  movel([0.304016, -1.350622, -2.573814, -0.787953, 1.570796, 1.874813],accel_mss,speed_ms,0,blend_radius_m)
  movel([0.304007, -1.350886, -2.573637, -0.787866, 1.570796, 1.874804],accel_mss,speed_ms,0,blend_radius_m)
  movel([0.303980, -1.351158, -2.573455, -0.787776, 1.570796, 1.874776],accel_mss,speed_ms,0,blend_radius_m)
  movel([0.303937, -1.351431, -2.573272, -0.787686, 1.570796, 1.874734],accel_mss,speed_ms,0,blend_radius_m)
  movel([0.303879, -1.351709, -2.573085, -0.787594, 1.570796, 1.874675],accel_mss,speed_ms,0,blend_radius_m)
  movel([0.303801, -1.351990, -2.572896, -0.787502, 1.570796, 1.874598],accel_mss,speed_ms,0,blend_radius_m)
  movel([0.303710, -1.352271, -2.572708, -0.787410, 1.570796, 1.874506],accel_mss,speed_ms,0,blend_radius_m)
  movel([0.303601, -1.352553, -2.572519, -0.787318, 1.570796, 1.874397],accel_mss,speed_ms,0,blend_radius_m)
  movel([0.303476, -1.352836, -2.572328, -0.787225, 1.570796, 1.874272],accel_mss,speed_ms,0,blend_radius_m)
  movel([0.303336, -1.353119, -2.572138, -0.787132, 1.570796, 1.874133],accel_mss,speed_ms,0,blend_radius_m)
  movel([0.303181, -1.353399, -2.571949, -0.787041, 1.570796, 1.873978],accel_mss,speed_ms,0,blend_radius_m)
  movel([0.303018, -1.353668, -2.571768, -0.786953, 1.570796, 1.873815],accel_mss,speed_ms,0,blend_radius_m)
  movel([0.302839, -1.353937, -2.571586, -0.786865, 1.570796, 1.873636],accel_mss,speed_ms,0,blend_radius_m)
  movel([0.302653, -1.354200, -2.571409, -0.786780, 1.570796, 1.873449],accel_mss,speed_ms,0,blend_radius_m)
  movel([0.302453, -1.354460, -2.571234, -0.786695, 1.570796, 1.873250],accel_mss,speed_ms,0,blend_radius_m)
  movel([0.302246, -1.354707, -2.571067, -0.786615, 1.570796, 1.873043],accel_mss,speed_ms,0,blend_radius_m)
  movel([0.302029, -1.354951, -2.570903, -0.786536, 1.570796, 1.872825],accel_mss,speed_ms,0,blend_radius_m)
  movel([0.301802, -1.355186, -2.570743, -0.786459, 1.570796, 1.872599],accel_mss,speed_ms,0,blend_radius_m)
  movel([0.301564, -1.355414, -2.570589, -0.786386, 1.570796, 1.872361],accel_mss,speed_ms,0,blend_radius_m)
  movel([0.301323, -1.355631, -2.570442, -0.786315, 1.570796, 1.872119],accel_mss,speed_ms,0,blend_radius_m)
  movel([0.301073, -1.355840, -2.570301, -0.786248, 1.570796, 1.871869],accel_mss,speed_ms,0,blend_radius_m)
  movel([0.300816, -1.356039, -2.570167, -0.786184, 1.570796, 1.871613],accel_mss,speed_ms,0,blend_radius_m)
  movel([0.300551, -1.356229, -2.570038, -0.786122, 1.570796, 1.871347],accel_mss,speed_ms,0,blend_radius_m)
  movel([0.300280, -1.356409, -2.569916, -0.786064, 1.570796, 1.871076],accel_mss,speed_ms,0,blend_radius_m)
  movel([0.300006, -1.356576, -2.569803, -0.786010, 1.570796, 1.870802],accel_mss,speed_ms,0,blend_radius_m)
  movel([0.299729, -1.356732, -2.569697, -0.785960, 1.570796, 1.870525],accel_mss,speed_ms,0,blend_radius_m)
  movel([0.299446, -1.356878, -2.569598, -0.785913, 1.570796, 1.870242],accel_mss,speed_ms,0,blend_radius_m)
  movel([0.299211, -1.356989, -2.569523, -0.785877, 1.570796, 1.870008],accel_mss,speed_ms,0,blend_radius_m)
  movel([0.298976, -1.357089, -2.569455, -0.785845, 1.570796, 1.869772],accel_mss,speed_ms,0,blend_radius_m)
  movel([0.298781, -1.357162, -2.569405, -0.785822, 1.570796, 1.869578],accel_mss,speed_ms,0,blend_radius_m)
  movel([0.298590, -1.357219, -2.569366, -0.785803, 1.570796, 1.869386],accel_mss,speed_ms,0,blend_radius_m)
  movel([0.298374, -1.357273, -2.569330, -0.785786, 1.570796, 1.869170],accel_mss,speed_ms,0,blend_radius_m)
  movel([0.298159, -1.357310, -2.569305, -0.785774, 1.570796, 1.868955],accel_mss,speed_ms,0,blend_radius_m)
  movel([0.297828, -1.357357, -2.569273, -0.785759, 1.570796, 1.868625],accel_mss,speed_ms,0,blend_radius_m)
  movel([0.297500, -1.357396, -2.569246, -0.785747, 1.570796, 1.868297],accel_mss,speed_ms,0,blend_radius_m)
  movel([0.297176, -1.357431, -2.569223, -0.785735, 1.570796, 1.867972],accel_mss,speed_ms,0,blend_radius_m)
  movel([0.296852, -1.357459, -2.569204, -0.785726, 1.570796, 1.867648],accel_mss,speed_ms,0,blend_radius_m)
  movel([0.296645, -1.357469, -2.569197, -0.785723, 1.570796, 1.867441],accel_mss,speed_ms,0,blend_radius_m)
  movel([0.296449, -1.357463, -2.569201, -0.785725, 1.570796, 1.867245],accel_mss,speed_ms,0,blend_radius_m)
  movel([0.296278, -1.357446, -2.569212, -0.785730, 1.570796, 1.867075],accel_mss,speed_ms,0,blend_radius_m)
  movel([0.296121, -1.357413, -2.569235, -0.785741, 1.570796, 1.866917],accel_mss,speed_ms,0,blend_radius_m)
  movel([0.295935, -1.357359, -2.569272, -0.785759, 1.570796, 1.866731],accel_mss,speed_ms,0,blend_radius_m)
  movel([0.295754, -1.357297, -2.569313, -0.785778, 1.570796, 1.866550],accel_mss,speed_ms,0,blend_radius_m)
  movel([0.295553, -1.357209, -2.569373, -0.785807, 1.570796, 1.866349],accel_mss,speed_ms,0,blend_radius_m)
  movel([0.295368, -1.357105, -2.569444, -0.785840, 1.570796, 1.866165],accel_mss,speed_ms,0,blend_radius_m)
  movel([0.295196, -1.356987, -2.569524, -0.785878, 1.570796, 1.865992],accel_mss,speed_ms,0,blend_radius_m)
  movel([0.295024, -1.356844, -2.569621, -0.785924, 1.570796, 1.865820],accel_mss,speed_ms,0,blend_radius_m)
  movel([0.294865, -1.356689, -2.569726, -0.785974, 1.570796, 1.865661],accel_mss,speed_ms,0,blend_radius_m)
  movel([0.294721, -1.356523, -2.569839, -0.786028, 1.570796, 1.865518],accel_mss,speed_ms,0,blend_radius_m)
  movel([0.294587, -1.356342, -2.569961, -0.786086, 1.570796, 1.865383],accel_mss,speed_ms,0,blend_radius_m)
  movel([0.294469, -1.356148, -2.570092, -0.786148, 1.570796, 1.865265],accel_mss,speed_ms,0,blend_radius_m)
  movel([0.294364, -1.355946, -2.570229, -0.786214, 1.570796, 1.865161],accel_mss,speed_ms,0,blend_radius_m)
  movel([0.294280, -1.355740, -2.570369, -0.786280, 1.570796, 1.865076],accel_mss,speed_ms,0,blend_radius_m)
  movel([0.294210, -1.355524, -2.570515, -0.786350, 1.570796, 1.865007],accel_mss,speed_ms,0,blend_radius_m)
  movel([0.294158, -1.355298, -2.570668, -0.786423, 1.570796, 1.864954],accel_mss,speed_ms,0,blend_radius_m)
  movel([0.294120, -1.355064, -2.570826, -0.786499, 1.570796, 1.864916],accel_mss,speed_ms,0,blend_radius_m)
  movel([0.294091, -1.354823, -2.570988, -0.786577, 1.570796, 1.864887],accel_mss,speed_ms,0,blend_radius_m)
  movel([0.294085, -1.354708, -2.571067, -0.786615, 1.570796, 1.864882],accel_mss,speed_ms,0,blend_radius_m)
  movel([0.294088, -1.354589, -2.571147, -0.786653, 1.570796, 1.864884],accel_mss,speed_ms,0,blend_radius_m)
  movel([0.294101, -1.354467, -2.571229, -0.786693, 1.570796, 1.864897],accel_mss,speed_ms,0,blend_radius_m)
  movel([0.294142, -1.354249, -2.571376, -0.786764, 1.570796, 1.864938],accel_mss,speed_ms,0,blend_radius_m)
  movel([0.294198, -1.354028, -2.571525, -0.786836, 1.570796, 1.864995],accel_mss,speed_ms,0,blend_radius_m)
  speed_ms = 0.003
  movel([0.294198, -1.341397, -2.565271, -0.805721, 1.570796, 1.864995],accel_mss,speed_ms,0,blend_radius_m)
  speed_ms = 0.01
  movel([0.294198, -1.317224, -2.552384, -0.842780, 1.570796, 1.864995],accel_mss,speed_ms,0,blend_radius_m)
  movel([0.288042, -1.339808, -2.537610, -0.834971, 1.570796, 1.858839],accel_mss,speed_ms,0,blend_radius_m)
  movel([0.288042, -1.363639, -2.550213, -0.798536, 1.570796, 1.858839],accel_mss,speed_ms,0,blend_radius_m)
  speed_ms = 0.003
  movel([0.288042, -1.372930, -2.554809, -0.784650, 1.570796, 1.858839],accel_mss,speed_ms,0,blend_radius_m)
  speed_ms = 0.007
  movel([0.288122, -1.372941, -2.554802, -0.784647, 1.570796, 1.858918],accel_mss,speed_ms,0,blend_radius_m)
  movel([0.288195, -1.372963, -2.554786, -0.784640, 1.570796, 1.858991],accel_mss,speed_ms,0,blend_radius_m)
  movel([0.288260, -1.372997, -2.554762, -0.784630, 1.570796, 1.859056],accel_mss,speed_ms,0,blend_radius_m)
  movel([0.288326, -1.373050, -2.554725, -0.784614, 1.570796, 1.859122],accel_mss,speed_ms,0,blend_radius_m)
  movel([0.288376, -1.373118, -2.554677, -0.784594, 1.570796, 1.859172],accel_mss,speed_ms,0,blend_radius_m)
  movel([0.288408, -1.373199, -2.554620, -0.784569, 1.570796, 1.859204],accel_mss,speed_ms,0,blend_radius_m)
  movel([0.288418, -1.373289, -2.554557, -0.784543, 1.570796, 1.859215],accel_mss,speed_ms,0,blend_radius_m)
  movel([0.288412, -1.373390, -2.554486, -0.784513, 1.570796, 1.859208],accel_mss,speed_ms,0,blend_radius_m)
  movel([0.288388, -1.373495, -2.554413, -0.784482, 1.570796, 1.859185],accel_mss,speed_ms,0,blend_radius_m)
  movel([0.288346, -1.373602, -2.554338, -0.784450, 1.570796, 1.859142],accel_mss,speed_ms,0,blend_radius_m)
  movel([0.288285, -1.373708, -2.554263, -0.784418, 1.570796, 1.859081],accel_mss,speed_ms,0,blend_radius_m)
  movel([0.288212, -1.373810, -2.554191, -0.784388, 1.570796, 1.859008],accel_mss,speed_ms,0,blend_radius_m)
  movel([0.288127, -1.373904, -2.554125, -0.784360, 1.570796, 1.858924],accel_mss,speed_ms,0,blend_radius_m)
  movel([0.288029, -1.373991, -2.554064, -0.784334, 1.570796, 1.858825],accel_mss,speed_ms,0,blend_radius_m)
  movel([0.287923, -1.374066, -2.554011, -0.784312, 1.570796, 1.858720],accel_mss,speed_ms,0,blend_radius_m)
  movel([0.287837, -1.374115, -2.553977, -0.784297, 1.570796, 1.858633],accel_mss,speed_ms,0,blend_radius_m)
  movel([0.287749, -1.374155, -2.553948, -0.784285, 1.570796, 1.858545],accel_mss,speed_ms,0,blend_radius_m)
  movel([0.287660, -1.374183, -2.553929, -0.784277, 1.570796, 1.858456],accel_mss,speed_ms,0,blend_radius_m)
  movel([0.287572, -1.374202, -2.553916, -0.784272, 1.570796, 1.858368],accel_mss,speed_ms,0,blend_radius_m)
  movel([0.287487, -1.374207, -2.553912, -0.784270, 1.570796, 1.858284],accel_mss,speed_ms,0,blend_radius_m)
  movel([0.287398, -1.374200, -2.553917, -0.784272, 1.570796, 1.858194],accel_mss,speed_ms,0,blend_radius_m)
  movel([0.287321, -1.374176, -2.553934, -0.784279, 1.570796, 1.858117],accel_mss,speed_ms,0,blend_radius_m)
  movel([0.287255, -1.374136, -2.553962, -0.784291, 1.570796, 1.858052],accel_mss,speed_ms,0,blend_radius_m)
  movel([0.287198, -1.374077, -2.554003, -0.784308, 1.570796, 1.857994],accel_mss,speed_ms,0,blend_radius_m)
  movel([0.287153, -1.374009, -2.554052, -0.784329, 1.570796, 1.857949],accel_mss,speed_ms,0,blend_radius_m)
  movel([0.287124, -1.373932, -2.554106, -0.784352, 1.570796, 1.857921],accel_mss,speed_ms,0,blend_radius_m)
  movel([0.287110, -1.373847, -2.554166, -0.784377, 1.570796, 1.857906],accel_mss,speed_ms,0,blend_radius_m)
  movel([0.287111, -1.373755, -2.554230, -0.784404, 1.570796, 1.857907],accel_mss,speed_ms,0,blend_radius_m)
  movel([0.287127, -1.373658, -2.554298, -0.784433, 1.570796, 1.857924],accel_mss,speed_ms,0,blend_radius_m)
  movel([0.287155, -1.373568, -2.554361, -0.784460, 1.570796, 1.857952],accel_mss,speed_ms,0,blend_radius_m)
  movel([0.287204, -1.373478, -2.554425, -0.784487, 1.570796, 1.858000],accel_mss,speed_ms,0,blend_radius_m)
  movel([0.287266, -1.373390, -2.554486, -0.784513, 1.570796, 1.858062],accel_mss,speed_ms,0,blend_radius_m)
  movel([0.287346, -1.373301, -2.554549, -0.784539, 1.570796, 1.858143],accel_mss,speed_ms,0,blend_radius_m)
  movel([0.287430, -1.373215, -2.554609, -0.784565, 1.570796, 1.858227],accel_mss,speed_ms,0,blend_radius_m)
  movel([0.287524, -1.373135, -2.554665, -0.784589, 1.570796, 1.858321],accel_mss,speed_ms,0,blend_radius_m)
  movel([0.287608, -1.373073, -2.554709, -0.784607, 1.570796, 1.858404],accel_mss,speed_ms,0,blend_radius_m)
  movel([0.287698, -1.373019, -2.554746, -0.784623, 1.570796, 1.858494],accel_mss,speed_ms,0,blend_radius_m)
  movel([0.287789, -1.372976, -2.554777, -0.784636, 1.570796, 1.858586],accel_mss,speed_ms,0,blend_radius_m)
  movel([0.287876, -1.372949, -2.554796, -0.784644, 1.570796, 1.858672],accel_mss,speed_ms,0,blend_radius_m)
  movel([0.287961, -1.372933, -2.554807, -0.784649, 1.570796, 1.858758],accel_mss,speed_ms,0,blend_radius_m)
  movel([0.288042, -1.372930, -2.554809, -0.784650, 1.570796, 1.858839],accel_mss,speed_ms,0,blend_radius_m)
  speed_ms = 0.003
  movel([0.288042, -1.376070, -2.556325, -0.779994, 1.570796, 1.858839],accel_mss,speed_ms,0,blend_radius_m)
  speed_ms = 0.007
  movel([0.288122, -1.376081, -2.556317, -0.779991, 1.570796, 1.858918],accel_mss,speed_ms,0,blend_radius_m)
  movel([0.288195, -1.376103, -2.556302, -0.779984, 1.570796, 1.858991],accel_mss,speed_ms,0,blend_radius_m)
  movel([0.288260, -1.376137, -2.556278, -0.779974, 1.570796, 1.859056],accel_mss,speed_ms,0,blend_radius_m)
  movel([0.288326, -1.376190, -2.556241, -0.779958, 1.570796, 1.859122],accel_mss,speed_ms,0,blend_radius_m)
  movel([0.288376, -1.376258, -2.556193, -0.779938, 1.570796, 1.859172],accel_mss,speed_ms,0,blend_radius_m)
  movel([0.288408, -1.376339, -2.556136, -0.779915, 1.570796, 1.859204],accel_mss,speed_ms,0,blend_radius_m)
  movel([0.288418, -1.376429, -2.556072, -0.779888, 1.570796, 1.859215],accel_mss,speed_ms,0,blend_radius_m)
  movel([0.288412, -1.376529, -2.556001, -0.779859, 1.570796, 1.859208],accel_mss,speed_ms,0,blend_radius_m)
  movel([0.288388, -1.376634, -2.555928, -0.779828, 1.570796, 1.859185],accel_mss,speed_ms,0,blend_radius_m)
  movel([0.288346, -1.376740, -2.555852, -0.779796, 1.570796, 1.859142],accel_mss,speed_ms,0,blend_radius_m)
  movel([0.288285, -1.376847, -2.555777, -0.779765, 1.570796, 1.859081],accel_mss,speed_ms,0,blend_radius_m)
  movel([0.288212, -1.376948, -2.555706, -0.779735, 1.570796, 1.859008],accel_mss,speed_ms,0,blend_radius_m)
  movel([0.288127, -1.377042, -2.555639, -0.779708, 1.570796, 1.858924],accel_mss,speed_ms,0,blend_radius_m)
  movel([0.288029, -1.377129, -2.555578, -0.779682, 1.570796, 1.858825],accel_mss,speed_ms,0,blend_radius_m)
  movel([0.287923, -1.377204, -2.555525, -0.779660, 1.570796, 1.858720],accel_mss,speed_ms,0,blend_radius_m)
  movel([0.287837, -1.377252, -2.555491, -0.779646, 1.570796, 1.858633],accel_mss,speed_ms,0,blend_radius_m)
  movel([0.287749, -1.377293, -2.555462, -0.779634, 1.570796, 1.858545],accel_mss,speed_ms,0,blend_radius_m)
  movel([0.287660, -1.377320, -2.555443, -0.779626, 1.570796, 1.858456],accel_mss,speed_ms,0,blend_radius_m)
  movel([0.287572, -1.377339, -2.555430, -0.779621, 1.570796, 1.858368],accel_mss,speed_ms,0,blend_radius_m)
  movel([0.287487, -1.377344, -2.555426, -0.779619, 1.570796, 1.858284],accel_mss,speed_ms,0,blend_radius_m)
  movel([0.287398, -1.377337, -2.555431, -0.779621, 1.570796, 1.858194],accel_mss,speed_ms,0,blend_radius_m)
  movel([0.287321, -1.377313, -2.555448, -0.779628, 1.570796, 1.858117],accel_mss,speed_ms,0,blend_radius_m)
  movel([0.287255, -1.377273, -2.555476, -0.779640, 1.570796, 1.858052],accel_mss,speed_ms,0,blend_radius_m)
  movel([0.287198, -1.377215, -2.555517, -0.779657, 1.570796, 1.857994],accel_mss,speed_ms,0,blend_radius_m)
  movel([0.287153, -1.377146, -2.555566, -0.779677, 1.570796, 1.857949],accel_mss,speed_ms,0,blend_radius_m)
  movel([0.287124, -1.377069, -2.555620, -0.779700, 1.570796, 1.857921],accel_mss,speed_ms,0,blend_radius_m)
  movel([0.287110, -1.376985, -2.555680, -0.779725, 1.570796, 1.857906],accel_mss,speed_ms,0,blend_radius_m)
  movel([0.287111, -1.376894, -2.555744, -0.779751, 1.570796, 1.857907],accel_mss,speed_ms,0,blend_radius_m)
  movel([0.287127, -1.376796, -2.555813, -0.779780, 1.570796, 1.857924],accel_mss,speed_ms,0,blend_radius_m)
  movel([0.287155, -1.376707, -2.555876, -0.779806, 1.570796, 1.857952],accel_mss,speed_ms,0,blend_radius_m)
  movel([0.287204, -1.376617, -2.555940, -0.779833, 1.570796, 1.858000],accel_mss,speed_ms,0,blend_radius_m)
  movel([0.287266, -1.376529, -2.556001, -0.779858, 1.570796, 1.858062],accel_mss,speed_ms,0,blend_radius_m)
  movel([0.287346, -1.376440, -2.556064, -0.779885, 1.570796, 1.858143],accel_mss,speed_ms,0,blend_radius_m)
  movel([0.287430, -1.376355, -2.556124, -0.779910, 1.570796, 1.858227],accel_mss,speed_ms,0,blend_radius_m)
  movel([0.287524, -1.376275, -2.556181, -0.779933, 1.570796, 1.858321],accel_mss,speed_ms,0,blend_radius_m)
  movel([0.287608, -1.376213, -2.556224, -0.779952, 1.570796, 1.858404],accel_mss,speed_ms,0,blend_radius_m)
  movel([0.287698, -1.376160, -2.556262, -0.779967, 1.570796, 1.858494],accel_mss,speed_ms,0,blend_radius_m)
  movel([0.287789, -1.376117, -2.556292, -0.779980, 1.570796, 1.858586],accel_mss,speed_ms,0,blend_radius_m)
  movel([0.287876, -1.376089, -2.556311, -0.779988, 1.570796, 1.858672],accel_mss,speed_ms,0,blend_radius_m)
  movel([0.287961, -1.376073, -2.556323, -0.779993, 1.570796, 1.858758],accel_mss,speed_ms,0,blend_radius_m)
  movel([0.288042, -1.376070, -2.556325, -0.779994, 1.570796, 1.858839],accel_mss,speed_ms,0,blend_radius_m)
  speed_ms = 0.003
  movel([0.288042, -1.363639, -2.550213, -0.798536, 1.570796, 1.858839],accel_mss,speed_ms,0,blend_radius_m)
  speed_ms = 0.01
  movel([0.288042, -1.339808, -2.537610, -0.834971, 1.570796, 1.858839],accel_mss,speed_ms,0,blend_radius_m)
  movel([0.266011, -1.335427, -2.540528, -0.836434, 1.570796, 1.836807],accel_mss,speed_ms,0,blend_radius_m)
  movel([0.266011, -1.359326, -2.553186, -0.799877, 1.570796, 1.836807],accel_mss,speed_ms,0,blend_radius_m)
  speed_ms = 0.003
  movel([0.266011, -1.368646, -2.557802, -0.785941, 1.570796, 1.836807],accel_mss,speed_ms,0,blend_radius_m)
  speed_ms = 0.007
  movel([0.265722, -1.369059, -2.557515, -0.785815, 1.570796, 1.836519],accel_mss,speed_ms,0,blend_radius_m)
  movel([0.265423, -1.369470, -2.557229, -0.785690, 1.570796, 1.836219],accel_mss,speed_ms,0,blend_radius_m)
  movel([0.265112, -1.369875, -2.556947, -0.785568, 1.570796, 1.835909],accel_mss,speed_ms,0,blend_radius_m)
  movel([0.264791, -1.370276, -2.556667, -0.785446, 1.570796, 1.835587],accel_mss,speed_ms,0,blend_radius_m)
  movel([0.264465, -1.370663, -2.556397, -0.785330, 1.570796, 1.835261],accel_mss,speed_ms,0,blend_radius_m)
  movel([0.264126, -1.371044, -2.556130, -0.785215, 1.570796, 1.834923],accel_mss,speed_ms,0,blend_radius_m)
  movel([0.263781, -1.371418, -2.555869, -0.785102, 1.570796, 1.834578],accel_mss,speed_ms,0,blend_radius_m)
  movel([0.263424, -1.371787, -2.555611, -0.784992, 1.570796, 1.834220],accel_mss,speed_ms,0,blend_radius_m)
  movel([0.263058, -1.372146, -2.555359, -0.784884, 1.570796, 1.833855],accel_mss,speed_ms,0,blend_radius_m)
  movel([0.262685, -1.372499, -2.555111, -0.784778, 1.570796, 1.833481],accel_mss,speed_ms,0,blend_radius_m)
  movel([0.262301, -1.372843, -2.554870, -0.784676, 1.570796, 1.833097],accel_mss,speed_ms,0,blend_radius_m)
  movel([0.261910, -1.373179, -2.554634, -0.784575, 1.570796, 1.832707],accel_mss,speed_ms,0,blend_radius_m)
  movel([0.261537, -1.373487, -2.554418, -0.784484, 1.570796, 1.832333],accel_mss,speed_ms,0,blend_radius_m)
  movel([0.261156, -1.373790, -2.554205, -0.784394, 1.570796, 1.831952],accel_mss,speed_ms,0,blend_radius_m)
  movel([0.260769, -1.374082, -2.554000, -0.784307, 1.570796, 1.831565],accel_mss,speed_ms,0,blend_radius_m)
  movel([0.260377, -1.374369, -2.553798, -0.784222, 1.570796, 1.831173],accel_mss,speed_ms,0,blend_radius_m)
  movel([0.259998, -1.374634, -2.553611, -0.784143, 1.570796, 1.830795],accel_mss,speed_ms,0,blend_radius_m)
  movel([0.259613, -1.374890, -2.553431, -0.784068, 1.570796, 1.830409],accel_mss,speed_ms,0,blend_radius_m)
  movel([0.259224, -1.375137, -2.553257, -0.783995, 1.570796, 1.830020],accel_mss,speed_ms,0,blend_radius_m)
  movel([0.258830, -1.375375, -2.553090, -0.783925, 1.570796, 1.829626],accel_mss,speed_ms,0,blend_radius_m)
  movel([0.258430, -1.375602, -2.552929, -0.783858, 1.570796, 1.829227],accel_mss,speed_ms,0,blend_radius_m)
  movel([0.258032, -1.375819, -2.552776, -0.783794, 1.570796, 1.828828],accel_mss,speed_ms,0,blend_radius_m)
  movel([0.257627, -1.376026, -2.552630, -0.783733, 1.570796, 1.828423],accel_mss,speed_ms,0,blend_radius_m)
  movel([0.257223, -1.376222, -2.552492, -0.783675, 1.570796, 1.828019],accel_mss,speed_ms,0,blend_radius_m)
  movel([0.256797, -1.376415, -2.552356, -0.783619, 1.570796, 1.827593],accel_mss,speed_ms,0,blend_radius_m)
  movel([0.256368, -1.376599, -2.552225, -0.783565, 1.570796, 1.827165],accel_mss,speed_ms,0,blend_radius_m)
  movel([0.255939, -1.376774, -2.552102, -0.783514, 1.570796, 1.826735],accel_mss,speed_ms,0,blend_radius_m)
  movel([0.255510, -1.376937, -2.551986, -0.783466, 1.570796, 1.826306],accel_mss,speed_ms,0,blend_radius_m)
  movel([0.255204, -1.377044, -2.551910, -0.783434, 1.570796, 1.826001],accel_mss,speed_ms,0,blend_radius_m)
  movel([0.254900, -1.377139, -2.551843, -0.783407, 1.570796, 1.825697],accel_mss,speed_ms,0,blend_radius_m)
  movel([0.254597, -1.377223, -2.551784, -0.783382, 1.570796, 1.825393],accel_mss,speed_ms,0,blend_radius_m)
  movel([0.254295, -1.377294, -2.551734, -0.783361, 1.570796, 1.825092],accel_mss,speed_ms,0,blend_radius_m)
  movel([0.253772, -1.377400, -2.551658, -0.783330, 1.570796, 1.824569],accel_mss,speed_ms,0,blend_radius_m)
  movel([0.253251, -1.377494, -2.551592, -0.783303, 1.570796, 1.824047],accel_mss,speed_ms,0,blend_radius_m)
  movel([0.252731, -1.377575, -2.551535, -0.783279, 1.570796, 1.823527],accel_mss,speed_ms,0,blend_radius_m)
  movel([0.252217, -1.377643, -2.551487, -0.783259, 1.570796, 1.823013],accel_mss,speed_ms,0,blend_radius_m)
  movel([0.251706, -1.377697, -2.551448, -0.783244, 1.570796, 1.822503],accel_mss,speed_ms,0,blend_radius_m)
  movel([0.251202, -1.377738, -2.551419, -0.783232, 1.570796, 1.821998],accel_mss,speed_ms,0,blend_radius_m)
  movel([0.250916, -1.377752, -2.551409, -0.783228, 1.570796, 1.821712],accel_mss,speed_ms,0,blend_radius_m)
  movel([0.250636, -1.377752, -2.551409, -0.783228, 1.570796, 1.821432],accel_mss,speed_ms,0,blend_radius_m)
  movel([0.250362, -1.377741, -2.551417, -0.783231, 1.570796, 1.821158],accel_mss,speed_ms,0,blend_radius_m)
  movel([0.250093, -1.377716, -2.551435, -0.783238, 1.570796, 1.820890],accel_mss,speed_ms,0,blend_radius_m)
  movel([0.249712, -1.377667, -2.551469, -0.783252, 1.570796, 1.820508],accel_mss,speed_ms,0,blend_radius_m)
  movel([0.249339, -1.377604, -2.551514, -0.783271, 1.570796, 1.820135],accel_mss,speed_ms,0,blend_radius_m)
  movel([0.248973, -1.377532, -2.551565, -0.783292, 1.570796, 1.819770],accel_mss,speed_ms,0,blend_radius_m)
  movel([0.248614, -1.377446, -2.551626, -0.783317, 1.570796, 1.819410],accel_mss,speed_ms,0,blend_radius_m)
  movel([0.248285, -1.377354, -2.551691, -0.783344, 1.570796, 1.819082],accel_mss,speed_ms,0,blend_radius_m)
  movel([0.247963, -1.377248, -2.551766, -0.783375, 1.570796, 1.818759],accel_mss,speed_ms,0,blend_radius_m)
  movel([0.247652, -1.377131, -2.551849, -0.783409, 1.570796, 1.818449],accel_mss,speed_ms,0,blend_radius_m)
  movel([0.247353, -1.376999, -2.551943, -0.783448, 1.570796, 1.818149],accel_mss,speed_ms,0,blend_radius_m)
  movel([0.247061, -1.376856, -2.552043, -0.783489, 1.570796, 1.817857],accel_mss,speed_ms,0,blend_radius_m)
  movel([0.246782, -1.376699, -2.552154, -0.783535, 1.570796, 1.817578],accel_mss,speed_ms,0,blend_radius_m)
  movel([0.246513, -1.376530, -2.552274, -0.783585, 1.570796, 1.817309],accel_mss,speed_ms,0,blend_radius_m)
  movel([0.246253, -1.376351, -2.552401, -0.783637, 1.570796, 1.817050],accel_mss,speed_ms,0,blend_radius_m)
  movel([0.245991, -1.376146, -2.552545, -0.783697, 1.570796, 1.816788],accel_mss,speed_ms,0,blend_radius_m)
  movel([0.245739, -1.375930, -2.552698, -0.783761, 1.570796, 1.816536],accel_mss,speed_ms,0,blend_radius_m)
  movel([0.245496, -1.375706, -2.552856, -0.783827, 1.570796, 1.816292],accel_mss,speed_ms,0,blend_radius_m)
  movel([0.245264, -1.375473, -2.553020, -0.783896, 1.570796, 1.816060],accel_mss,speed_ms,0,blend_radius_m)
  movel([0.245040, -1.375220, -2.553198, -0.783970, 1.570796, 1.815836],accel_mss,speed_ms,0,blend_radius_m)
  movel([0.244827, -1.374957, -2.553384, -0.784048, 1.570796, 1.815624],accel_mss,speed_ms,0,blend_radius_m)
  movel([0.244629, -1.374686, -2.553575, -0.784128, 1.570796, 1.815425],accel_mss,speed_ms,0,blend_radius_m)
  movel([0.244442, -1.374403, -2.553774, -0.784212, 1.570796, 1.815238],accel_mss,speed_ms,0,blend_radius_m)
  movel([0.244275, -1.374114, -2.553978, -0.784298, 1.570796, 1.815071],accel_mss,speed_ms,0,blend_radius_m)
  movel([0.244119, -1.373818, -2.554185, -0.784385, 1.570796, 1.814915],accel_mss,speed_ms,0,blend_radius_m)
  movel([0.243980, -1.373509, -2.554403, -0.784477, 1.570796, 1.814777],accel_mss,speed_ms,0,blend_radius_m)
  movel([0.243857, -1.373194, -2.554624, -0.784571, 1.570796, 1.814654],accel_mss,speed_ms,0,blend_radius_m)
  movel([0.243743, -1.372861, -2.554857, -0.784670, 1.570796, 1.814539],accel_mss,speed_ms,0,blend_radius_m)
  movel([0.243647, -1.372520, -2.555097, -0.784772, 1.570796, 1.814444],accel_mss,speed_ms,0,blend_radius_m)
  movel([0.243565, -1.372169, -2.555343, -0.784877, 1.570796, 1.814362],accel_mss,speed_ms,0,blend_radius_m)
  movel([0.243497, -1.371812, -2.555593, -0.784984, 1.570796, 1.814293],accel_mss,speed_ms,0,blend_radius_m)
  movel([0.243441, -1.371423, -2.555865, -0.785101, 1.570796, 1.814237],accel_mss,speed_ms,0,blend_radius_m)
  movel([0.243401, -1.371029, -2.556141, -0.785219, 1.570796, 1.814197],accel_mss,speed_ms,0,blend_radius_m)
  movel([0.243370, -1.370631, -2.556418, -0.785339, 1.570796, 1.814167],accel_mss,speed_ms,0,blend_radius_m)
  movel([0.243356, -1.370224, -2.556703, -0.785462, 1.570796, 1.814152],accel_mss,speed_ms,0,blend_radius_m)
  movel([0.243358, -1.369940, -2.556901, -0.785548, 1.570796, 1.814154],accel_mss,speed_ms,0,blend_radius_m)
  movel([0.243372, -1.369653, -2.557101, -0.785635, 1.570796, 1.814168],accel_mss,speed_ms,0,blend_radius_m)
  movel([0.243400, -1.369383, -2.557289, -0.785717, 1.570796, 1.814196],accel_mss,speed_ms,0,blend_radius_m)
  movel([0.243440, -1.369110, -2.557480, -0.785800, 1.570796, 1.814237],accel_mss,speed_ms,0,blend_radius_m)
  movel([0.243512, -1.368755, -2.557726, -0.785907, 1.570796, 1.814308],accel_mss,speed_ms,0,blend_radius_m)
  movel([0.243598, -1.368399, -2.557975, -0.786016, 1.570796, 1.814394],accel_mss,speed_ms,0,blend_radius_m)
  movel([0.243753, -1.367791, -2.558397, -0.786201, 1.570796, 1.814549],accel_mss,speed_ms,0,blend_radius_m)
  movel([0.243913, -1.367182, -2.558820, -0.786387, 1.570796, 1.814710],accel_mss,speed_ms,0,blend_radius_m)
  movel([0.244088, -1.366544, -2.559262, -0.786583, 1.570796, 1.814885],accel_mss,speed_ms,0,blend_radius_m)
  movel([0.244266, -1.365905, -2.559704, -0.786780, 1.570796, 1.815063],accel_mss,speed_ms,0,blend_radius_m)
  movel([0.244375, -1.365550, -2.559950, -0.786889, 1.570796, 1.815172],accel_mss,speed_ms,0,blend_radius_m)
  movel([0.244496, -1.365193, -2.560197, -0.787000, 1.570796, 1.815293],accel_mss,speed_ms,0,blend_radius_m)
  movel([0.244610, -1.364899, -2.560399, -0.787090, 1.570796, 1.815406],accel_mss,speed_ms,0,blend_radius_m)
  movel([0.244742, -1.364607, -2.560601, -0.787181, 1.570796, 1.815538],accel_mss,speed_ms,0,blend_radius_m)
  movel([0.244917, -1.364247, -2.560849, -0.787292, 1.570796, 1.815713],accel_mss,speed_ms,0,blend_radius_m)
  movel([0.245104, -1.363888, -2.561097, -0.787404, 1.570796, 1.815901],accel_mss,speed_ms,0,blend_radius_m)
  movel([0.245373, -1.363400, -2.561433, -0.787556, 1.570796, 1.816169],accel_mss,speed_ms,0,blend_radius_m)
  movel([0.245657, -1.362916, -2.561766, -0.787707, 1.570796, 1.816453],accel_mss,speed_ms,0,blend_radius_m)
  movel([0.245957, -1.362433, -2.562098, -0.787858, 1.570796, 1.816753],accel_mss,speed_ms,0,blend_radius_m)
  movel([0.246272, -1.361954, -2.562427, -0.788008, 1.570796, 1.817069],accel_mss,speed_ms,0,blend_radius_m)
  movel([0.246604, -1.361477, -2.562754, -0.788158, 1.570796, 1.817400],accel_mss,speed_ms,0,blend_radius_m)
  movel([0.246948, -1.361006, -2.563077, -0.788306, 1.570796, 1.817745],accel_mss,speed_ms,0,blend_radius_m)
  movel([0.247308, -1.360539, -2.563397, -0.788453, 1.570796, 1.818104],accel_mss,speed_ms,0,blend_radius_m)
  movel([0.247669, -1.360096, -2.563700, -0.788593, 1.570796, 1.818465],accel_mss,speed_ms,0,blend_radius_m)
  movel([0.248045, -1.359657, -2.564001, -0.788732, 1.570796, 1.818841],accel_mss,speed_ms,0,blend_radius_m)
  movel([0.248433, -1.359226, -2.564295, -0.788868, 1.570796, 1.819229],accel_mss,speed_ms,0,blend_radius_m)
  movel([0.248835, -1.358804, -2.564583, -0.789002, 1.570796, 1.819632],accel_mss,speed_ms,0,blend_radius_m)
  movel([0.249250, -1.358389, -2.564866, -0.789135, 1.570796, 1.820047],accel_mss,speed_ms,0,blend_radius_m)
  movel([0.249677, -1.357985, -2.565141, -0.789263, 1.570796, 1.820473],accel_mss,speed_ms,0,blend_radius_m)
  movel([0.250113, -1.357588, -2.565411, -0.789390, 1.570796, 1.820909],accel_mss,speed_ms,0,blend_radius_m)
  movel([0.250553, -1.357212, -2.565667, -0.789510, 1.570796, 1.821349],accel_mss,speed_ms,0,blend_radius_m)
  movel([0.251003, -1.356845, -2.565916, -0.789628, 1.570796, 1.821799],accel_mss,speed_ms,0,blend_radius_m)
  movel([0.251461, -1.356491, -2.566157, -0.789741, 1.570796, 1.822257],accel_mss,speed_ms,0,blend_radius_m)
  movel([0.251928, -1.356150, -2.566388, -0.789851, 1.570796, 1.822724],accel_mss,speed_ms,0,blend_radius_m)
  movel([0.252401, -1.355820, -2.566612, -0.789957, 1.570796, 1.823197],accel_mss,speed_ms,0,blend_radius_m)
  movel([0.252882, -1.355506, -2.566825, -0.790058, 1.570796, 1.823678],accel_mss,speed_ms,0,blend_radius_m)
  movel([0.253371, -1.355203, -2.567030, -0.790156, 1.570796, 1.824168],accel_mss,speed_ms,0,blend_radius_m)
  movel([0.253864, -1.354916, -2.567224, -0.790249, 1.570796, 1.824661],accel_mss,speed_ms,0,blend_radius_m)
  movel([0.254363, -1.354644, -2.567408, -0.790337, 1.570796, 1.825159],accel_mss,speed_ms,0,blend_radius_m)
  movel([0.254864, -1.354386, -2.567583, -0.790420, 1.570796, 1.825660],accel_mss,speed_ms,0,blend_radius_m)
  movel([0.255371, -1.354143, -2.567747, -0.790499, 1.570796, 1.826167],accel_mss,speed_ms,0,blend_radius_m)
  movel([0.255878, -1.353918, -2.567899, -0.790572, 1.570796, 1.826674],accel_mss,speed_ms,0,blend_radius_m)
  movel([0.256388, -1.353708, -2.568041, -0.790640, 1.570796, 1.827184],accel_mss,speed_ms,0,blend_radius_m)
  movel([0.256897, -1.353516, -2.568170, -0.790703, 1.570796, 1.827694],accel_mss,speed_ms,0,blend_radius_m)
  movel([0.257220, -1.353405, -2.568245, -0.790739, 1.570796, 1.828016],accel_mss,speed_ms,0,blend_radius_m)
  movel([0.257542, -1.353304, -2.568314, -0.790772, 1.570796, 1.828339],accel_mss,speed_ms,0,blend_radius_m)
  movel([0.257864, -1.353213, -2.568375, -0.790801, 1.570796, 1.828660],accel_mss,speed_ms,0,blend_radius_m)
  movel([0.258186, -1.353132, -2.568430, -0.790828, 1.570796, 1.828982],accel_mss,speed_ms,0,blend_radius_m)
  movel([0.258674, -1.353025, -2.568501, -0.790863, 1.570796, 1.829471],accel_mss,speed_ms,0,blend_radius_m)
  movel([0.259162, -1.352930, -2.568565, -0.790894, 1.570796, 1.829958],accel_mss,speed_ms,0,blend_radius_m)
  movel([0.259643, -1.352852, -2.568618, -0.790919, 1.570796, 1.830439],accel_mss,speed_ms,0,blend_radius_m)
  movel([0.260122, -1.352787, -2.568662, -0.790940, 1.570796, 1.830918],accel_mss,speed_ms,0,blend_radius_m)
  movel([0.260597, -1.352739, -2.568694, -0.790956, 1.570796, 1.831393],accel_mss,speed_ms,0,blend_radius_m)
  movel([0.261066, -1.352703, -2.568719, -0.790968, 1.570796, 1.831862],accel_mss,speed_ms,0,blend_radius_m)
  movel([0.261368, -1.352691, -2.568726, -0.790971, 1.570796, 1.832164],accel_mss,speed_ms,0,blend_radius_m)
  movel([0.261664, -1.352690, -2.568727, -0.790972, 1.570796, 1.832461],accel_mss,speed_ms,0,blend_radius_m)
  movel([0.261955, -1.352700, -2.568720, -0.790969, 1.570796, 1.832752],accel_mss,speed_ms,0,blend_radius_m)
  movel([0.262241, -1.352720, -2.568707, -0.790962, 1.570796, 1.833038],accel_mss,speed_ms,0,blend_radius_m)
  movel([0.262661, -1.352767, -2.568675, -0.790947, 1.570796, 1.833457],accel_mss,speed_ms,0,blend_radius_m)
  movel([0.263068, -1.352832, -2.568631, -0.790925, 1.570796, 1.833864],accel_mss,speed_ms,0,blend_radius_m)
  movel([0.263465, -1.352914, -2.568576, -0.790899, 1.570796, 1.834261],accel_mss,speed_ms,0,blend_radius_m)
  movel([0.263854, -1.353010, -2.568511, -0.790867, 1.570796, 1.834650],accel_mss,speed_ms,0,blend_radius_m)
  movel([0.264230, -1.353124, -2.568434, -0.790830, 1.570796, 1.835026],accel_mss,speed_ms,0,blend_radius_m)
  movel([0.264596, -1.353255, -2.568346, -0.790788, 1.570796, 1.835393],accel_mss,speed_ms,0,blend_radius_m)
  movel([0.264949, -1.353402, -2.568247, -0.790740, 1.570796, 1.835745],accel_mss,speed_ms,0,blend_radius_m)
  movel([0.265290, -1.353563, -2.568138, -0.790687, 1.570796, 1.836086],accel_mss,speed_ms,0,blend_radius_m)
  movel([0.265619, -1.353742, -2.568017, -0.790629, 1.570796, 1.836415],accel_mss,speed_ms,0,blend_radius_m)
  movel([0.265932, -1.353935, -2.567888, -0.790567, 1.570796, 1.836728],accel_mss,speed_ms,0,blend_radius_m)
  movel([0.266233, -1.354144, -2.567746, -0.790499, 1.570796, 1.837029],accel_mss,speed_ms,0,blend_radius_m)
  movel([0.266520, -1.354367, -2.567596, -0.790427, 1.570796, 1.837317],accel_mss,speed_ms,0,blend_radius_m)
  movel([0.266792, -1.354605, -2.567434, -0.790349, 1.570796, 1.837588],accel_mss,speed_ms,0,blend_radius_m)
  movel([0.267049, -1.354857, -2.567264, -0.790268, 1.570796, 1.837846],accel_mss,speed_ms,0,blend_radius_m)
  movel([0.267289, -1.355121, -2.567085, -0.790182, 1.570796, 1.838085],accel_mss,speed_ms,0,blend_radius_m)
  movel([0.267517, -1.355401, -2.566896, -0.790092, 1.570796, 1.838314],accel_mss,speed_ms,0,blend_radius_m)
  movel([0.267728, -1.355692, -2.566698, -0.789998, 1.570796, 1.838524],accel_mss,speed_ms,0,blend_radius_m)
  movel([0.267923, -1.355997, -2.566492, -0.789900, 1.570796, 1.838719],accel_mss,speed_ms,0,blend_radius_m)
  movel([0.268100, -1.356312, -2.566278, -0.789799, 1.570796, 1.838896],accel_mss,speed_ms,0,blend_radius_m)
  movel([0.268259, -1.356641, -2.566055, -0.789693, 1.570796, 1.839056],accel_mss,speed_ms,0,blend_radius_m)
  movel([0.268402, -1.356970, -2.565831, -0.789588, 1.570796, 1.839199],accel_mss,speed_ms,0,blend_radius_m)
  movel([0.268531, -1.357306, -2.565603, -0.789480, 1.570796, 1.839328],accel_mss,speed_ms,0,blend_radius_m)
  movel([0.268646, -1.357649, -2.565369, -0.789370, 1.570796, 1.839442],accel_mss,speed_ms,0,blend_radius_m)
  movel([0.268740, -1.357976, -2.565147, -0.789266, 1.570796, 1.839536],accel_mss,speed_ms,0,blend_radius_m)
  movel([0.268817, -1.358311, -2.564918, -0.789159, 1.570796, 1.839614],accel_mss,speed_ms,0,blend_radius_m)
  movel([0.268879, -1.358653, -2.564685, -0.789050, 1.570796, 1.839675],accel_mss,speed_ms,0,blend_radius_m)
  movel([0.268926, -1.359012, -2.564440, -0.788936, 1.570796, 1.839722],accel_mss,speed_ms,0,blend_radius_m)
  movel([0.268959, -1.359378, -2.564191, -0.788820, 1.570796, 1.839755],accel_mss,speed_ms,0,blend_radius_m)
  movel([0.268974, -1.359750, -2.563937, -0.788702, 1.570796, 1.839770],accel_mss,speed_ms,0,blend_radius_m)
  movel([0.268978, -1.360174, -2.563647, -0.788568, 1.570796, 1.839774],accel_mss,speed_ms,0,blend_radius_m)
  movel([0.268967, -1.360604, -2.563353, -0.788433, 1.570796, 1.839763],accel_mss,speed_ms,0,blend_radius_m)
  movel([0.268945, -1.361035, -2.563057, -0.788297, 1.570796, 1.839742],accel_mss,speed_ms,0,blend_radius_m)
  movel([0.268920, -1.361344, -2.562846, -0.788200, 1.570796, 1.839717],accel_mss,speed_ms,0,blend_radius_m)
  movel([0.268878, -1.361657, -2.562631, -0.788101, 1.570796, 1.839674],accel_mss,speed_ms,0,blend_radius_m)
  movel([0.268822, -1.361974, -2.562414, -0.788002, 1.570796, 1.839619],accel_mss,speed_ms,0,blend_radius_m)
  movel([0.268755, -1.362292, -2.562195, -0.787902, 1.570796, 1.839551],accel_mss,speed_ms,0,blend_radius_m)
  movel([0.268618, -1.362832, -2.561824, -0.787733, 1.570796, 1.839414],accel_mss,speed_ms,0,blend_radius_m)
  movel([0.268469, -1.363376, -2.561450, -0.787563, 1.570796, 1.839265],accel_mss,speed_ms,0,blend_radius_m)
  movel([0.268302, -1.363921, -2.561074, -0.787394, 1.570796, 1.839099],accel_mss,speed_ms,0,blend_radius_m)
  movel([0.268119, -1.364471, -2.560695, -0.787223, 1.570796, 1.838915],accel_mss,speed_ms,0,blend_radius_m)
  movel([0.267921, -1.365022, -2.560315, -0.787052, 1.570796, 1.838717],accel_mss,speed_ms,0,blend_radius_m)
  movel([0.267709, -1.365572, -2.559934, -0.786882, 1.570796, 1.838506],accel_mss,speed_ms,0,blend_radius_m)
  movel([0.267571, -1.365903, -2.559706, -0.786780, 1.570796, 1.838368],accel_mss,speed_ms,0,blend_radius_m)
  movel([0.267421, -1.366235, -2.559476, -0.786678, 1.570796, 1.838218],accel_mss,speed_ms,0,blend_radius_m)
  movel([0.267258, -1.366567, -2.559246, -0.786576, 1.570796, 1.838054],accel_mss,speed_ms,0,blend_radius_m)
  movel([0.267080, -1.366898, -2.559016, -0.786474, 1.570796, 1.837877],accel_mss,speed_ms,0,blend_radius_m)
  movel([0.266832, -1.367339, -2.558711, -0.786339, 1.570796, 1.837628],accel_mss,speed_ms,0,blend_radius_m)
  movel([0.266570, -1.367777, -2.558407, -0.786206, 1.570796, 1.837367],accel_mss,speed_ms,0,blend_radius_m)
  movel([0.266296, -1.368212, -2.558104, -0.786073, 1.570796, 1.837092],accel_mss,speed_ms,0,blend_radius_m)
  movel([0.266011, -1.368646, -2.557802, -0.785941, 1.570796, 1.836807],accel_mss,speed_ms,0,blend_radius_m)
  speed_ms = 0.003
  movel([0.266011, -1.371796, -2.559325, -0.781267, 1.570796, 1.836807],accel_mss,speed_ms,0,blend_radius_m)
  speed_ms = 0.007
  movel([0.265722, -1.372208, -2.559037, -0.781144, 1.570796, 1.836519],accel_mss,speed_ms,0,blend_radius_m)
  movel([0.265423, -1.372619, -2.558750, -0.781020, 1.570796, 1.836219],accel_mss,speed_ms,0,blend_radius_m)
  movel([0.265112, -1.373022, -2.558467, -0.780899, 1.570796, 1.835909],accel_mss,speed_ms,0,blend_radius_m)
  movel([0.264791, -1.373423, -2.558187, -0.780780, 1.570796, 1.835587],accel_mss,speed_ms,0,blend_radius_m)
  movel([0.264465, -1.373808, -2.557916, -0.780665, 1.570796, 1.835261],accel_mss,speed_ms,0,blend_radius_m)
  movel([0.264126, -1.374189, -2.557649, -0.780551, 1.570796, 1.834923],accel_mss,speed_ms,0,blend_radius_m)
  movel([0.263781, -1.374562, -2.557387, -0.780440, 1.570796, 1.834578],accel_mss,speed_ms,0,blend_radius_m)
  movel([0.263424, -1.374930, -2.557128, -0.780331, 1.570796, 1.834220],accel_mss,speed_ms,0,blend_radius_m)
  movel([0.263058, -1.375288, -2.556876, -0.780225, 1.570796, 1.833855],accel_mss,speed_ms,0,blend_radius_m)
  movel([0.262685, -1.375640, -2.556628, -0.780121, 1.570796, 1.833481],accel_mss,speed_ms,0,blend_radius_m)
  movel([0.262301, -1.375984, -2.556386, -0.780019, 1.570796, 1.833097],accel_mss,speed_ms,0,blend_radius_m)
  movel([0.261910, -1.376319, -2.556150, -0.779920, 1.570796, 1.832707],accel_mss,speed_ms,0,blend_radius_m)
  movel([0.261537, -1.376626, -2.555933, -0.779830, 1.570796, 1.832333],accel_mss,speed_ms,0,blend_radius_m)
  movel([0.261156, -1.376928, -2.555720, -0.779741, 1.570796, 1.831952],accel_mss,speed_ms,0,blend_radius_m)
  movel([0.260769, -1.377220, -2.555514, -0.779656, 1.570796, 1.831565],accel_mss,speed_ms,0,blend_radius_m)
  movel([0.260377, -1.377506, -2.555312, -0.779572, 1.570796, 1.831173],accel_mss,speed_ms,0,blend_radius_m)
  movel([0.259998, -1.377770, -2.555124, -0.779494, 1.570796, 1.830795],accel_mss,speed_ms,0,blend_radius_m)
  movel([0.259613, -1.378025, -2.554944, -0.779420, 1.570796, 1.830409],accel_mss,speed_ms,0,blend_radius_m)
  movel([0.259224, -1.378272, -2.554769, -0.779348, 1.570796, 1.830020],accel_mss,speed_ms,0,blend_radius_m)
  movel([0.258830, -1.378509, -2.554601, -0.779278, 1.570796, 1.829626],accel_mss,speed_ms,0,blend_radius_m)
  movel([0.258430, -1.378736, -2.554441, -0.779212, 1.570796, 1.829227],accel_mss,speed_ms,0,blend_radius_m)
  movel([0.258032, -1.378952, -2.554287, -0.779149, 1.570796, 1.828828],accel_mss,speed_ms,0,blend_radius_m)
  movel([0.257627, -1.379159, -2.554141, -0.779089, 1.570796, 1.828423],accel_mss,speed_ms,0,blend_radius_m)
  movel([0.257223, -1.379354, -2.554002, -0.779033, 1.570796, 1.828019],accel_mss,speed_ms,0,blend_radius_m)
  movel([0.256797, -1.379547, -2.553866, -0.778977, 1.570796, 1.827593],accel_mss,speed_ms,0,blend_radius_m)
  movel([0.256368, -1.379731, -2.553735, -0.778923, 1.570796, 1.827165],accel_mss,speed_ms,0,blend_radius_m)
  movel([0.255939, -1.379905, -2.553612, -0.778873, 1.570796, 1.826735],accel_mss,speed_ms,0,blend_radius_m)
  movel([0.255510, -1.380068, -2.553496, -0.778826, 1.570796, 1.826306],accel_mss,speed_ms,0,blend_radius_m)
  movel([0.255204, -1.380175, -2.553419, -0.778795, 1.570796, 1.826001],accel_mss,speed_ms,0,blend_radius_m)
  movel([0.254900, -1.380269, -2.553352, -0.778767, 1.570796, 1.825697],accel_mss,speed_ms,0,blend_radius_m)
  movel([0.254597, -1.380353, -2.553293, -0.778743, 1.570796, 1.825393],accel_mss,speed_ms,0,blend_radius_m)
  movel([0.254295, -1.380423, -2.553243, -0.778723, 1.570796, 1.825092],accel_mss,speed_ms,0,blend_radius_m)
  movel([0.253772, -1.380530, -2.553167, -0.778692, 1.570796, 1.824569],accel_mss,speed_ms,0,blend_radius_m)
  movel([0.253251, -1.380623, -2.553100, -0.778665, 1.570796, 1.824047],accel_mss,speed_ms,0,blend_radius_m)
  movel([0.252731, -1.380704, -2.553043, -0.778642, 1.570796, 1.823527],accel_mss,speed_ms,0,blend_radius_m)
  movel([0.252217, -1.380772, -2.552995, -0.778622, 1.570796, 1.823013],accel_mss,speed_ms,0,blend_radius_m)
  movel([0.251706, -1.380826, -2.552956, -0.778607, 1.570796, 1.822503],accel_mss,speed_ms,0,blend_radius_m)
  movel([0.251202, -1.380867, -2.552927, -0.778595, 1.570796, 1.821998],accel_mss,speed_ms,0,blend_radius_m)
  movel([0.250916, -1.380881, -2.552917, -0.778591, 1.570796, 1.821712],accel_mss,speed_ms,0,blend_radius_m)
  movel([0.250636, -1.380881, -2.552917, -0.778591, 1.570796, 1.821432],accel_mss,speed_ms,0,blend_radius_m)
  movel([0.250362, -1.380870, -2.552925, -0.778594, 1.570796, 1.821158],accel_mss,speed_ms,0,blend_radius_m)
  movel([0.250093, -1.380845, -2.552943, -0.778601, 1.570796, 1.820890],accel_mss,speed_ms,0,blend_radius_m)
  movel([0.249712, -1.380796, -2.552978, -0.778615, 1.570796, 1.820508],accel_mss,speed_ms,0,blend_radius_m)
  movel([0.249339, -1.380733, -2.553022, -0.778633, 1.570796, 1.820135],accel_mss,speed_ms,0,blend_radius_m)
  movel([0.248973, -1.380661, -2.553073, -0.778654, 1.570796, 1.819770],accel_mss,speed_ms,0,blend_radius_m)
  movel([0.248614, -1.380576, -2.553134, -0.778679, 1.570796, 1.819410],accel_mss,speed_ms,0,blend_radius_m)
  movel([0.248285, -1.380483, -2.553200, -0.778706, 1.570796, 1.819082],accel_mss,speed_ms,0,blend_radius_m)
  movel([0.247963, -1.380378, -2.553275, -0.778736, 1.570796, 1.818759],accel_mss,speed_ms,0,blend_radius_m)
  movel([0.247652, -1.380262, -2.553358, -0.778770, 1.570796, 1.818449],accel_mss,speed_ms,0,blend_radius_m)
  movel([0.247353, -1.380129, -2.553452, -0.778808, 1.570796, 1.818149],accel_mss,speed_ms,0,blend_radius_m)
  movel([0.247061, -1.379987, -2.553553, -0.778849, 1.570796, 1.817857],accel_mss,speed_ms,0,blend_radius_m)
  movel([0.246782, -1.379830, -2.553664, -0.778894, 1.570796, 1.817578],accel_mss,speed_ms,0,blend_radius_m)
  movel([0.246513, -1.379662, -2.553784, -0.778943, 1.570796, 1.817309],accel_mss,speed_ms,0,blend_radius_m)
  movel([0.246253, -1.379483, -2.553911, -0.778995, 1.570796, 1.817050],accel_mss,speed_ms,0,blend_radius_m)
  movel([0.245991, -1.379279, -2.554056, -0.779054, 1.570796, 1.816788],accel_mss,speed_ms,0,blend_radius_m)
  movel([0.245739, -1.379063, -2.554209, -0.779117, 1.570796, 1.816536],accel_mss,speed_ms,0,blend_radius_m)
  movel([0.245496, -1.378839, -2.554367, -0.779182, 1.570796, 1.816292],accel_mss,speed_ms,0,blend_radius_m)
  movel([0.245264, -1.378607, -2.554532, -0.779250, 1.570796, 1.816060],accel_mss,speed_ms,0,blend_radius_m)
  movel([0.245040, -1.378355, -2.554710, -0.779323, 1.570796, 1.815836],accel_mss,speed_ms,0,blend_radius_m)
  movel([0.244827, -1.378093, -2.554896, -0.779400, 1.570796, 1.815624],accel_mss,speed_ms,0,blend_radius_m)
  movel([0.244629, -1.377822, -2.555088, -0.779479, 1.570796, 1.815425],accel_mss,speed_ms,0,blend_radius_m)
  movel([0.244442, -1.377540, -2.555287, -0.779562, 1.570796, 1.815238],accel_mss,speed_ms,0,blend_radius_m)
  movel([0.244275, -1.377251, -2.555491, -0.779646, 1.570796, 1.815071],accel_mss,speed_ms,0,blend_radius_m)
  movel([0.244119, -1.376956, -2.555700, -0.779733, 1.570796, 1.814915],accel_mss,speed_ms,0,blend_radius_m)
  movel([0.243980, -1.376648, -2.555917, -0.779824, 1.570796, 1.814777],accel_mss,speed_ms,0,blend_radius_m)
  movel([0.243857, -1.376333, -2.556140, -0.779916, 1.570796, 1.814654],accel_mss,speed_ms,0,blend_radius_m)
  movel([0.243743, -1.376002, -2.556373, -0.780014, 1.570796, 1.814539],accel_mss,speed_ms,0,blend_radius_m)
  movel([0.243647, -1.375661, -2.556614, -0.780115, 1.570796, 1.814444],accel_mss,speed_ms,0,blend_radius_m)
  movel([0.243565, -1.375311, -2.556860, -0.780218, 1.570796, 1.814362],accel_mss,speed_ms,0,blend_radius_m)
  movel([0.243497, -1.374955, -2.557110, -0.780324, 1.570796, 1.814293],accel_mss,speed_ms,0,blend_radius_m)
  movel([0.243441, -1.374567, -2.557383, -0.780439, 1.570796, 1.814237],accel_mss,speed_ms,0,blend_radius_m)
  movel([0.243401, -1.374174, -2.557659, -0.780556, 1.570796, 1.814197],accel_mss,speed_ms,0,blend_radius_m)
  movel([0.243370, -1.373777, -2.557938, -0.780674, 1.570796, 1.814167],accel_mss,speed_ms,0,blend_radius_m)
  movel([0.243356, -1.373371, -2.558223, -0.780795, 1.570796, 1.814152],accel_mss,speed_ms,0,blend_radius_m)
  movel([0.243358, -1.373087, -2.558422, -0.780880, 1.570796, 1.814154],accel_mss,speed_ms,0,blend_radius_m)
  movel([0.243372, -1.372801, -2.558622, -0.780966, 1.570796, 1.814168],accel_mss,speed_ms,0,blend_radius_m)
  movel([0.243400, -1.372532, -2.558811, -0.781046, 1.570796, 1.814196],accel_mss,speed_ms,0,blend_radius_m)
  movel([0.243440, -1.372259, -2.559002, -0.781128, 1.570796, 1.814237],accel_mss,speed_ms,0,blend_radius_m)
  movel([0.243512, -1.371905, -2.559249, -0.781235, 1.570796, 1.814308],accel_mss,speed_ms,0,blend_radius_m)
  movel([0.243598, -1.371550, -2.559498, -0.781342, 1.570796, 1.814394],accel_mss,speed_ms,0,blend_radius_m)
  movel([0.243753, -1.370943, -2.559921, -0.781525, 1.570796, 1.814549],accel_mss,speed_ms,0,blend_radius_m)
  movel([0.243913, -1.370336, -2.560345, -0.781709, 1.570796, 1.814710],accel_mss,speed_ms,0,blend_radius_m)
  movel([0.244088, -1.369700, -2.560788, -0.781902, 1.570796, 1.814885],accel_mss,speed_ms,0,blend_radius_m)
  movel([0.244266, -1.369062, -2.561231, -0.782096, 1.570796, 1.815063],accel_mss,speed_ms,0,blend_radius_m)
  movel([0.244375, -1.368708, -2.561477, -0.782204, 1.570796, 1.815172],accel_mss,speed_ms,0,blend_radius_m)
  movel([0.244496, -1.368351, -2.561725, -0.782313, 1.570796, 1.815293],accel_mss,speed_ms,0,blend_radius_m)
  movel([0.244610, -1.368059, -2.561928, -0.782402, 1.570796, 1.815406],accel_mss,speed_ms,0,blend_radius_m)
  movel([0.244742, -1.367767, -2.562130, -0.782492, 1.570796, 1.815538],accel_mss,speed_ms,0,blend_radius_m)
  movel([0.244917, -1.367408, -2.562379, -0.782602, 1.570796, 1.815713],accel_mss,speed_ms,0,blend_radius_m)
  movel([0.245104, -1.367049, -2.562627, -0.782712, 1.570796, 1.815901],accel_mss,speed_ms,0,blend_radius_m)
  movel([0.245373, -1.366563, -2.562964, -0.782862, 1.570796, 1.816169],accel_mss,speed_ms,0,blend_radius_m)
  movel([0.245657, -1.366080, -2.563298, -0.783011, 1.570796, 1.816453],accel_mss,speed_ms,0,blend_radius_m)
  movel([0.245957, -1.365598, -2.563631, -0.783160, 1.570796, 1.816753],accel_mss,speed_ms,0,blend_radius_m)
  movel([0.246272, -1.365120, -2.563960, -0.783308, 1.570796, 1.817069],accel_mss,speed_ms,0,blend_radius_m)
  movel([0.246604, -1.364644, -2.564289, -0.783456, 1.570796, 1.817400],accel_mss,speed_ms,0,blend_radius_m)
  movel([0.246948, -1.364175, -2.564612, -0.783602, 1.570796, 1.817745],accel_mss,speed_ms,0,blend_radius_m)
  movel([0.247308, -1.363709, -2.564933, -0.783748, 1.570796, 1.818104],accel_mss,speed_ms,0,blend_radius_m)
  movel([0.247669, -1.363267, -2.565237, -0.783886, 1.570796, 1.818465],accel_mss,speed_ms,0,blend_radius_m)
  movel([0.248045, -1.362828, -2.565538, -0.784023, 1.570796, 1.818841],accel_mss,speed_ms,0,blend_radius_m)
  movel([0.248433, -1.362399, -2.565832, -0.784158, 1.570796, 1.819229],accel_mss,speed_ms,0,blend_radius_m)
  movel([0.248835, -1.361978, -2.566121, -0.784290, 1.570796, 1.819632],accel_mss,speed_ms,0,blend_radius_m)
  movel([0.249250, -1.361563, -2.566405, -0.784421, 1.570796, 1.820047],accel_mss,speed_ms,0,blend_radius_m)
  movel([0.249677, -1.361160, -2.566681, -0.784548, 1.570796, 1.820473],accel_mss,speed_ms,0,blend_radius_m)
  movel([0.250113, -1.360764, -2.566952, -0.784673, 1.570796, 1.820909],accel_mss,speed_ms,0,blend_radius_m)
  movel([0.250553, -1.360389, -2.567208, -0.784792, 1.570796, 1.821349],accel_mss,speed_ms,0,blend_radius_m)
  movel([0.251003, -1.360024, -2.567457, -0.784908, 1.570796, 1.821799],accel_mss,speed_ms,0,blend_radius_m)
  movel([0.251461, -1.359670, -2.567699, -0.785020, 1.570796, 1.822257],accel_mss,speed_ms,0,blend_radius_m)
  movel([0.251928, -1.359330, -2.567930, -0.785128, 1.570796, 1.822724],accel_mss,speed_ms,0,blend_radius_m)
  movel([0.252401, -1.359000, -2.568155, -0.785233, 1.570796, 1.823197],accel_mss,speed_ms,0,blend_radius_m)
  movel([0.252882, -1.358687, -2.568369, -0.785333, 1.570796, 1.823678],accel_mss,speed_ms,0,blend_radius_m)
  movel([0.253371, -1.358385, -2.568574, -0.785430, 1.570796, 1.824168],accel_mss,speed_ms,0,blend_radius_m)
  movel([0.253864, -1.358099, -2.568769, -0.785521, 1.570796, 1.824661],accel_mss,speed_ms,0,blend_radius_m)
  movel([0.254363, -1.357827, -2.568954, -0.785608, 1.570796, 1.825159],accel_mss,speed_ms,0,blend_radius_m)
  movel([0.254864, -1.357570, -2.569128, -0.785691, 1.570796, 1.825660],accel_mss,speed_ms,0,blend_radius_m)
  movel([0.255371, -1.357328, -2.569293, -0.785769, 1.570796, 1.826167],accel_mss,speed_ms,0,blend_radius_m)
  movel([0.255878, -1.357103, -2.569445, -0.785841, 1.570796, 1.826674],accel_mss,speed_ms,0,blend_radius_m)
  movel([0.256388, -1.356894, -2.569587, -0.785908, 1.570796, 1.827184],accel_mss,speed_ms,0,blend_radius_m)
  movel([0.256897, -1.356702, -2.569717, -0.785970, 1.570796, 1.827694],accel_mss,speed_ms,0,blend_radius_m)
  movel([0.257220, -1.356592, -2.569792, -0.786005, 1.570796, 1.828016],accel_mss,speed_ms,0,blend_radius_m)
  movel([0.257542, -1.356490, -2.569861, -0.786038, 1.570796, 1.828339],accel_mss,speed_ms,0,blend_radius_m)
  movel([0.257864, -1.356400, -2.569922, -0.786067, 1.570796, 1.828660],accel_mss,speed_ms,0,blend_radius_m)
  movel([0.258186, -1.356318, -2.569977, -0.786093, 1.570796, 1.828982],accel_mss,speed_ms,0,blend_radius_m)
  movel([0.258674, -1.356212, -2.570049, -0.786128, 1.570796, 1.829471],accel_mss,speed_ms,0,blend_radius_m)
  movel([0.259162, -1.356117, -2.570113, -0.786158, 1.570796, 1.829958],accel_mss,speed_ms,0,blend_radius_m)
  movel([0.259643, -1.356039, -2.570166, -0.786184, 1.570796, 1.830439],accel_mss,speed_ms,0,blend_radius_m)
  movel([0.260122, -1.355975, -2.570210, -0.786204, 1.570796, 1.830918],accel_mss,speed_ms,0,blend_radius_m)
  movel([0.260597, -1.355926, -2.570243, -0.786220, 1.570796, 1.831393],accel_mss,speed_ms,0,blend_radius_m)
  movel([0.261066, -1.355890, -2.570267, -0.786232, 1.570796, 1.831862],accel_mss,speed_ms,0,blend_radius_m)
  movel([0.261368, -1.355879, -2.570275, -0.786235, 1.570796, 1.832164],accel_mss,speed_ms,0,blend_radius_m)
  movel([0.261664, -1.355877, -2.570276, -0.786236, 1.570796, 1.832461],accel_mss,speed_ms,0,blend_radius_m)
  movel([0.261955, -1.355888, -2.570269, -0.786232, 1.570796, 1.832752],accel_mss,speed_ms,0,blend_radius_m)
  movel([0.262241, -1.355908, -2.570255, -0.786226, 1.570796, 1.833038],accel_mss,speed_ms,0,blend_radius_m)
  movel([0.262661, -1.355955, -2.570223, -0.786211, 1.570796, 1.833457],accel_mss,speed_ms,0,blend_radius_m)
  movel([0.263068, -1.356020, -2.570180, -0.786190, 1.570796, 1.833864],accel_mss,speed_ms,0,blend_radius_m)
  movel([0.263465, -1.356101, -2.570124, -0.786163, 1.570796, 1.834261],accel_mss,speed_ms,0,blend_radius_m)
  movel([0.263854, -1.356197, -2.570059, -0.786132, 1.570796, 1.834650],accel_mss,speed_ms,0,blend_radius_m)
  movel([0.264230, -1.356311, -2.569982, -0.786096, 1.570796, 1.835026],accel_mss,speed_ms,0,blend_radius_m)
  movel([0.264596, -1.356442, -2.569894, -0.786054, 1.570796, 1.835393],accel_mss,speed_ms,0,blend_radius_m)
  movel([0.264949, -1.356588, -2.569794, -0.786006, 1.570796, 1.835745],accel_mss,speed_ms,0,blend_radius_m)
  movel([0.265290, -1.356749, -2.569685, -0.785955, 1.570796, 1.836086],accel_mss,speed_ms,0,blend_radius_m)
  movel([0.265619, -1.356928, -2.569564, -0.785897, 1.570796, 1.836415],accel_mss,speed_ms,0,blend_radius_m)
  movel([0.265932, -1.357120, -2.569434, -0.785835, 1.570796, 1.836728],accel_mss,speed_ms,0,blend_radius_m)
  movel([0.266233, -1.357329, -2.569292, -0.785768, 1.570796, 1.837029],accel_mss,speed_ms,0,blend_radius_m)
  movel([0.266520, -1.357551, -2.569141, -0.785697, 1.570796, 1.837317],accel_mss,speed_ms,0,blend_radius_m)
  movel([0.266792, -1.357789, -2.568980, -0.785621, 1.570796, 1.837588],accel_mss,speed_ms,0,blend_radius_m)
  movel([0.267049, -1.358039, -2.568809, -0.785540, 1.570796, 1.837846],accel_mss,speed_ms,0,blend_radius_m)
  movel([0.267289, -1.358304, -2.568630, -0.785456, 1.570796, 1.838085],accel_mss,speed_ms,0,blend_radius_m)
  movel([0.267517, -1.358583, -2.568440, -0.785367, 1.570796, 1.838314],accel_mss,speed_ms,0,blend_radius_m)
  movel([0.267728, -1.358873, -2.568242, -0.785274, 1.570796, 1.838524],accel_mss,speed_ms,0,blend_radius_m)
  movel([0.267923, -1.359177, -2.568035, -0.785177, 1.570796, 1.838719],accel_mss,speed_ms,0,blend_radius_m)
  movel([0.268100, -1.359492, -2.567820, -0.785077, 1.570796, 1.838896],accel_mss,speed_ms,0,blend_radius_m)
  movel([0.268259, -1.359820, -2.567596, -0.784973, 1.570796, 1.839056],accel_mss,speed_ms,0,blend_radius_m)
  movel([0.268402, -1.360148, -2.567372, -0.784868, 1.570796, 1.839199],accel_mss,speed_ms,0,blend_radius_m)
  movel([0.268531, -1.360483, -2.567144, -0.784762, 1.570796, 1.839328],accel_mss,speed_ms,0,blend_radius_m)
  movel([0.268646, -1.360826, -2.566910, -0.784654, 1.570796, 1.839442],accel_mss,speed_ms,0,blend_radius_m)
  movel([0.268740, -1.361151, -2.566687, -0.784551, 1.570796, 1.839536],accel_mss,speed_ms,0,blend_radius_m)
  movel([0.268817, -1.361486, -2.566458, -0.784445, 1.570796, 1.839614],accel_mss,speed_ms,0,blend_radius_m)
  movel([0.268879, -1.361827, -2.566224, -0.784338, 1.570796, 1.839675],accel_mss,speed_ms,0,blend_radius_m)
  movel([0.268926, -1.362186, -2.565979, -0.784225, 1.570796, 1.839722],accel_mss,speed_ms,0,blend_radius_m)
  movel([0.268959, -1.362550, -2.565729, -0.784110, 1.570796, 1.839755],accel_mss,speed_ms,0,blend_radius_m)
  movel([0.268974, -1.362921, -2.565474, -0.783994, 1.570796, 1.839770],accel_mss,speed_ms,0,blend_radius_m)
  movel([0.268978, -1.363344, -2.565183, -0.783862, 1.570796, 1.839774],accel_mss,speed_ms,0,blend_radius_m)
  movel([0.268967, -1.363773, -2.564888, -0.783727, 1.570796, 1.839763],accel_mss,speed_ms,0,blend_radius_m)
  movel([0.268945, -1.364203, -2.564592, -0.783593, 1.570796, 1.839742],accel_mss,speed_ms,0,blend_radius_m)
  movel([0.268920, -1.364511, -2.564380, -0.783497, 1.570796, 1.839717],accel_mss,speed_ms,0,blend_radius_m)
  movel([0.268878, -1.364824, -2.564165, -0.783400, 1.570796, 1.839674],accel_mss,speed_ms,0,blend_radius_m)
  movel([0.268822, -1.365140, -2.563947, -0.783302, 1.570796, 1.839619],accel_mss,speed_ms,0,blend_radius_m)
  movel([0.268755, -1.365457, -2.563728, -0.783204, 1.570796, 1.839551],accel_mss,speed_ms,0,blend_radius_m)
  movel([0.268618, -1.365996, -2.563356, -0.783037, 1.570796, 1.839414],accel_mss,speed_ms,0,blend_radius_m)
  movel([0.268469, -1.366539, -2.562981, -0.782869, 1.570796, 1.839265],accel_mss,speed_ms,0,blend_radius_m)
  movel([0.268302, -1.367083, -2.562604, -0.782702, 1.570796, 1.839099],accel_mss,speed_ms,0,blend_radius_m)
  movel([0.268119, -1.367631, -2.562224, -0.782533, 1.570796, 1.838915],accel_mss,speed_ms,0,blend_radius_m)
  movel([0.267921, -1.368181, -2.561843, -0.782365, 1.570796, 1.838717],accel_mss,speed_ms,0,blend_radius_m)
  movel([0.267709, -1.368730, -2.561462, -0.782197, 1.570796, 1.838506],accel_mss,speed_ms,0,blend_radius_m)
  movel([0.267571, -1.369060, -2.561233, -0.782096, 1.570796, 1.838368],accel_mss,speed_ms,0,blend_radius_m)
  movel([0.267421, -1.369391, -2.561002, -0.781995, 1.570796, 1.838218],accel_mss,speed_ms,0,blend_radius_m)
  movel([0.267258, -1.369722, -2.560772, -0.781895, 1.570796, 1.838054],accel_mss,speed_ms,0,blend_radius_m)
  movel([0.267080, -1.370053, -2.560542, -0.781794, 1.570796, 1.837877],accel_mss,speed_ms,0,blend_radius_m)
  movel([0.266832, -1.370492, -2.560235, -0.781661, 1.570796, 1.837628],accel_mss,speed_ms,0,blend_radius_m)
  movel([0.266570, -1.370929, -2.559931, -0.781529, 1.570796, 1.837367],accel_mss,speed_ms,0,blend_radius_m)
  movel([0.266296, -1.371363, -2.559628, -0.781398, 1.570796, 1.837092],accel_mss,speed_ms,0,blend_radius_m)
  movel([0.266011, -1.371796, -2.559325, -0.781267, 1.570796, 1.836807],accel_mss,speed_ms,0,blend_radius_m)
  speed_ms = 0.003
  movel([0.266011, -1.359326, -2.553186, -0.799877, 1.570796, 1.836807],accel_mss,speed_ms,0,blend_radius_m)
  speed_ms = 0.01
  movel([0.266011, -1.335427, -2.540528, -0.836434, 1.570796, 1.836807],accel_mss,speed_ms,0,blend_radius_m)
  movel([0.264726, -1.335140, -2.540718, -0.836531, 1.570796, 1.835522],accel_mss,speed_ms,0,blend_radius_m)
  movel([0.264726, -1.359043, -2.553380, -0.799966, 1.570796, 1.835522],accel_mss,speed_ms,0,blend_radius_m)
  speed_ms = 0.003
  movel([0.264726, -1.368365, -2.557998, -0.786026, 1.570796, 1.835522],accel_mss,speed_ms,0,blend_radius_m)
  speed_ms = 0.007
  movel([0.264459, -1.368745, -2.557734, -0.785910, 1.570796, 1.835255],accel_mss,speed_ms,0,blend_radius_m)
  movel([0.264181, -1.369124, -2.557470, -0.785795, 1.570796, 1.834978],accel_mss,speed_ms,0,blend_radius_m)
  movel([0.263892, -1.369495, -2.557211, -0.785683, 1.570796, 1.834688],accel_mss,speed_ms,0,blend_radius_m)
  movel([0.263592, -1.369864, -2.556954, -0.785571, 1.570796, 1.834388],accel_mss,speed_ms,0,blend_radius_m)
  movel([0.263283, -1.370225, -2.556702, -0.785462, 1.570796, 1.834079],accel_mss,speed_ms,0,blend_radius_m)
  movel([0.262963, -1.370583, -2.556452, -0.785354, 1.570796, 1.833759],accel_mss,speed_ms,0,blend_radius_m)
  movel([0.262632, -1.370934, -2.556207, -0.785248, 1.570796, 1.833428],accel_mss,speed_ms,0,blend_radius_m)
  movel([0.262300, -1.371271, -2.555971, -0.785146, 1.570796, 1.833096],accel_mss,speed_ms,0,blend_radius_m)
  movel([0.261959, -1.371602, -2.555740, -0.785047, 1.570796, 1.832755],accel_mss,speed_ms,0,blend_radius_m)
  movel([0.261608, -1.371924, -2.555514, -0.784950, 1.570796, 1.832404],accel_mss,speed_ms,0,blend_radius_m)
  movel([0.261251, -1.372239, -2.555294, -0.784856, 1.570796, 1.832047],accel_mss,speed_ms,0,blend_radius_m)
  movel([0.260885, -1.372547, -2.555078, -0.784764, 1.570796, 1.831681],accel_mss,speed_ms,0,blend_radius_m)
  movel([0.260512, -1.372845, -2.554869, -0.784675, 1.570796, 1.831308],accel_mss,speed_ms,0,blend_radius_m)
  movel([0.260133, -1.373134, -2.554666, -0.784589, 1.570796, 1.830929],accel_mss,speed_ms,0,blend_radius_m)
  movel([0.259752, -1.373411, -2.554471, -0.784506, 1.570796, 1.830549],accel_mss,speed_ms,0,blend_radius_m)
  movel([0.259369, -1.373676, -2.554285, -0.784428, 1.570796, 1.830165],accel_mss,speed_ms,0,blend_radius_m)
  movel([0.258979, -1.373933, -2.554105, -0.784351, 1.570796, 1.829775],accel_mss,speed_ms,0,blend_radius_m)
  movel([0.258583, -1.374178, -2.553933, -0.784279, 1.570796, 1.829379],accel_mss,speed_ms,0,blend_radius_m)
  movel([0.258183, -1.374412, -2.553768, -0.784209, 1.570796, 1.828979],accel_mss,speed_ms,0,blend_radius_m)
  movel([0.257780, -1.374634, -2.553611, -0.784143, 1.570796, 1.828576],accel_mss,speed_ms,0,blend_radius_m)
  movel([0.257376, -1.374846, -2.553462, -0.784081, 1.570796, 1.828172],accel_mss,speed_ms,0,blend_radius_m)
  movel([0.256961, -1.375046, -2.553321, -0.784022, 1.570796, 1.827757],accel_mss,speed_ms,0,blend_radius_m)
  movel([0.256546, -1.375232, -2.553191, -0.783967, 1.570796, 1.827342],accel_mss,speed_ms,0,blend_radius_m)
  movel([0.256128, -1.375402, -2.553070, -0.783917, 1.570796, 1.826924],accel_mss,speed_ms,0,blend_radius_m)
  movel([0.255708, -1.375556, -2.552962, -0.783871, 1.570796, 1.826504],accel_mss,speed_ms,0,blend_radius_m)
  movel([0.255290, -1.375695, -2.552864, -0.783830, 1.570796, 1.826086],accel_mss,speed_ms,0,blend_radius_m)
  movel([0.254850, -1.375824, -2.552772, -0.783792, 1.570796, 1.825646],accel_mss,speed_ms,0,blend_radius_m)
  movel([0.254411, -1.375938, -2.552692, -0.783759, 1.570796, 1.825208],accel_mss,speed_ms,0,blend_radius_m)
  movel([0.253975, -1.376037, -2.552622, -0.783730, 1.570796, 1.824771],accel_mss,speed_ms,0,blend_radius_m)
  movel([0.253540, -1.376123, -2.552561, -0.783704, 1.570796, 1.824336],accel_mss,speed_ms,0,blend_radius_m)
  movel([0.253112, -1.376191, -2.552513, -0.783684, 1.570796, 1.823908],accel_mss,speed_ms,0,blend_radius_m)
  movel([0.252686, -1.376244, -2.552476, -0.783669, 1.570796, 1.823483],accel_mss,speed_ms,0,blend_radius_m)
  movel([0.252264, -1.376284, -2.552448, -0.783657, 1.570796, 1.823061],accel_mss,speed_ms,0,blend_radius_m)
  movel([0.251849, -1.376305, -2.552433, -0.783651, 1.570796, 1.822646],accel_mss,speed_ms,0,blend_radius_m)
  movel([0.251441, -1.376314, -2.552427, -0.783648, 1.570796, 1.822237],accel_mss,speed_ms,0,blend_radius_m)
  movel([0.251039, -1.376304, -2.552434, -0.783651, 1.570796, 1.821835],accel_mss,speed_ms,0,blend_radius_m)
  movel([0.250665, -1.376279, -2.552451, -0.783659, 1.570796, 1.821461],accel_mss,speed_ms,0,blend_radius_m)
  movel([0.250299, -1.376238, -2.552480, -0.783671, 1.570796, 1.821095],accel_mss,speed_ms,0,blend_radius_m)
  movel([0.249945, -1.376179, -2.552522, -0.783688, 1.570796, 1.820742],accel_mss,speed_ms,0,blend_radius_m)
  movel([0.249601, -1.376103, -2.552575, -0.783710, 1.570796, 1.820397],accel_mss,speed_ms,0,blend_radius_m)
  movel([0.249268, -1.376009, -2.552642, -0.783738, 1.570796, 1.820064],accel_mss,speed_ms,0,blend_radius_m)
  movel([0.248923, -1.375893, -2.552724, -0.783772, 1.570796, 1.819719],accel_mss,speed_ms,0,blend_radius_m)
  movel([0.248591, -1.375760, -2.552818, -0.783811, 1.570796, 1.819387],accel_mss,speed_ms,0,blend_radius_m)
  movel([0.248271, -1.375611, -2.552923, -0.783855, 1.570796, 1.819067],accel_mss,speed_ms,0,blend_radius_m)
  movel([0.247963, -1.375447, -2.553039, -0.783903, 1.570796, 1.818760],accel_mss,speed_ms,0,blend_radius_m)
  movel([0.247671, -1.375267, -2.553165, -0.783956, 1.570796, 1.818468],accel_mss,speed_ms,0,blend_radius_m)
  movel([0.247393, -1.375074, -2.553302, -0.784014, 1.570796, 1.818189],accel_mss,speed_ms,0,blend_radius_m)
  movel([0.247127, -1.374865, -2.553449, -0.784075, 1.570796, 1.817923],accel_mss,speed_ms,0,blend_radius_m)
  movel([0.246876, -1.374643, -2.553605, -0.784141, 1.570796, 1.817673],accel_mss,speed_ms,0,blend_radius_m)
  movel([0.246644, -1.374404, -2.553774, -0.784212, 1.570796, 1.817440],accel_mss,speed_ms,0,blend_radius_m)
  movel([0.246416, -1.374146, -2.553955, -0.784288, 1.570796, 1.817213],accel_mss,speed_ms,0,blend_radius_m)
  movel([0.246206, -1.373876, -2.554145, -0.784368, 1.570796, 1.817002],accel_mss,speed_ms,0,blend_radius_m)
  movel([0.246010, -1.373594, -2.554343, -0.784452, 1.570796, 1.816806],accel_mss,speed_ms,0,blend_radius_m)
  movel([0.245831, -1.373300, -2.554550, -0.784540, 1.570796, 1.816628],accel_mss,speed_ms,0,blend_radius_m)
  movel([0.245667, -1.372994, -2.554764, -0.784631, 1.570796, 1.816463],accel_mss,speed_ms,0,blend_radius_m)
  movel([0.245521, -1.372677, -2.554987, -0.784725, 1.570796, 1.816318],accel_mss,speed_ms,0,blend_radius_m)
  movel([0.245390, -1.372351, -2.555215, -0.784823, 1.570796, 1.816186],accel_mss,speed_ms,0,blend_radius_m)
  movel([0.245275, -1.372014, -2.555452, -0.784924, 1.570796, 1.816071],accel_mss,speed_ms,0,blend_radius_m)
  movel([0.245179, -1.371667, -2.555694, -0.785028, 1.570796, 1.815975],accel_mss,speed_ms,0,blend_radius_m)
  movel([0.245098, -1.371305, -2.555947, -0.785136, 1.570796, 1.815894],accel_mss,speed_ms,0,blend_radius_m)
  movel([0.245033, -1.370936, -2.556205, -0.785247, 1.570796, 1.815829],accel_mss,speed_ms,0,blend_radius_m)
  movel([0.244986, -1.370558, -2.556470, -0.785361, 1.570796, 1.815783],accel_mss,speed_ms,0,blend_radius_m)
  movel([0.244956, -1.370173, -2.556739, -0.785478, 1.570796, 1.815752],accel_mss,speed_ms,0,blend_radius_m)
  movel([0.244943, -1.369780, -2.557012, -0.785596, 1.570796, 1.815739],accel_mss,speed_ms,0,blend_radius_m)
  movel([0.244948, -1.369380, -2.557291, -0.785717, 1.570796, 1.815745],accel_mss,speed_ms,0,blend_radius_m)
  movel([0.244971, -1.368975, -2.557573, -0.785840, 1.570796, 1.815768],accel_mss,speed_ms,0,blend_radius_m)
  movel([0.245012, -1.368563, -2.557860, -0.785966, 1.570796, 1.815809],accel_mss,speed_ms,0,blend_radius_m)
  movel([0.245068, -1.368148, -2.558149, -0.786092, 1.570796, 1.815864],accel_mss,speed_ms,0,blend_radius_m)
  movel([0.245143, -1.367730, -2.558439, -0.786220, 1.570796, 1.815940],accel_mss,speed_ms,0,blend_radius_m)
  movel([0.245235, -1.367309, -2.558731, -0.786349, 1.570796, 1.816032],accel_mss,speed_ms,0,blend_radius_m)
  movel([0.245345, -1.366885, -2.559025, -0.786478, 1.570796, 1.816141],accel_mss,speed_ms,0,blend_radius_m)
  movel([0.245471, -1.366456, -2.559323, -0.786610, 1.570796, 1.816268],accel_mss,speed_ms,0,blend_radius_m)
  movel([0.245615, -1.366027, -2.559620, -0.786742, 1.570796, 1.816411],accel_mss,speed_ms,0,blend_radius_m)
  movel([0.245777, -1.365596, -2.559918, -0.786875, 1.570796, 1.816573],accel_mss,speed_ms,0,blend_radius_m)
  movel([0.245954, -1.365165, -2.560216, -0.787008, 1.570796, 1.816750],accel_mss,speed_ms,0,blend_radius_m)
  movel([0.246150, -1.364730, -2.560516, -0.787143, 1.570796, 1.816946],accel_mss,speed_ms,0,blend_radius_m)
  movel([0.246359, -1.364298, -2.560814, -0.787277, 1.570796, 1.817156],accel_mss,speed_ms,0,blend_radius_m)
  movel([0.246577, -1.363879, -2.561103, -0.787407, 1.570796, 1.817373],accel_mss,speed_ms,0,blend_radius_m)
  movel([0.246806, -1.363461, -2.561391, -0.787537, 1.570796, 1.817603],accel_mss,speed_ms,0,blend_radius_m)
  movel([0.247047, -1.363045, -2.561678, -0.787667, 1.570796, 1.817843],accel_mss,speed_ms,0,blend_radius_m)
  movel([0.247299, -1.362629, -2.561964, -0.787797, 1.570796, 1.818095],accel_mss,speed_ms,0,blend_radius_m)
  movel([0.247538, -1.362256, -2.562220, -0.787913, 1.570796, 1.818334],accel_mss,speed_ms,0,blend_radius_m)
  movel([0.247791, -1.361887, -2.562473, -0.788029, 1.570796, 1.818588],accel_mss,speed_ms,0,blend_radius_m)
  movel([0.248054, -1.361521, -2.562724, -0.788144, 1.570796, 1.818850],accel_mss,speed_ms,0,blend_radius_m)
  movel([0.248331, -1.361162, -2.562971, -0.788257, 1.570796, 1.819128],accel_mss,speed_ms,0,blend_radius_m)
  movel([0.248616, -1.360809, -2.563212, -0.788368, 1.570796, 1.819412],accel_mss,speed_ms,0,blend_radius_m)
  movel([0.248911, -1.360462, -2.563450, -0.788477, 1.570796, 1.819708],accel_mss,speed_ms,0,blend_radius_m)
  movel([0.249219, -1.360121, -2.563683, -0.788585, 1.570796, 1.820015],accel_mss,speed_ms,0,blend_radius_m)
  movel([0.249537, -1.359788, -2.563911, -0.788690, 1.570796, 1.820333],accel_mss,speed_ms,0,blend_radius_m)
  movel([0.249891, -1.359433, -2.564153, -0.788803, 1.570796, 1.820687],accel_mss,speed_ms,0,blend_radius_m)
  movel([0.250253, -1.359084, -2.564392, -0.788914, 1.570796, 1.821049],accel_mss,speed_ms,0,blend_radius_m)
  movel([0.250622, -1.358742, -2.564625, -0.789022, 1.570796, 1.821419],accel_mss,speed_ms,0,blend_radius_m)
  movel([0.251000, -1.358407, -2.564853, -0.789129, 1.570796, 1.821796],accel_mss,speed_ms,0,blend_radius_m)
  movel([0.251409, -1.358057, -2.565092, -0.789240, 1.570796, 1.822206],accel_mss,speed_ms,0,blend_radius_m)
  movel([0.251825, -1.357718, -2.565322, -0.789348, 1.570796, 1.822622],accel_mss,speed_ms,0,blend_radius_m)
  movel([0.252250, -1.357385, -2.565549, -0.789455, 1.570796, 1.823046],accel_mss,speed_ms,0,blend_radius_m)
  movel([0.252636, -1.357097, -2.565745, -0.789547, 1.570796, 1.823432],accel_mss,speed_ms,0,blend_radius_m)
  movel([0.253029, -1.356819, -2.565934, -0.789636, 1.570796, 1.823825],accel_mss,speed_ms,0,blend_radius_m)
  movel([0.253428, -1.356554, -2.566114, -0.789721, 1.570796, 1.824225],accel_mss,speed_ms,0,blend_radius_m)
  movel([0.253830, -1.356305, -2.566283, -0.789801, 1.570796, 1.824626],accel_mss,speed_ms,0,blend_radius_m)
  movel([0.254233, -1.356070, -2.566442, -0.789877, 1.570796, 1.825029],accel_mss,speed_ms,0,blend_radius_m)
  movel([0.254642, -1.355847, -2.566594, -0.789949, 1.570796, 1.825438],accel_mss,speed_ms,0,blend_radius_m)
  movel([0.255090, -1.355620, -2.566747, -0.790022, 1.570796, 1.825886],accel_mss,speed_ms,0,blend_radius_m)
  movel([0.255537, -1.355405, -2.566893, -0.790091, 1.570796, 1.826333],accel_mss,speed_ms,0,blend_radius_m)
  movel([0.255988, -1.355202, -2.567031, -0.790157, 1.570796, 1.826784],accel_mss,speed_ms,0,blend_radius_m)
  movel([0.256396, -1.355028, -2.567149, -0.790213, 1.570796, 1.827192],accel_mss,speed_ms,0,blend_radius_m)
  movel([0.256803, -1.354865, -2.567259, -0.790265, 1.570796, 1.827599],accel_mss,speed_ms,0,blend_radius_m)
  movel([0.256987, -1.354795, -2.567306, -0.790288, 1.570796, 1.827783],accel_mss,speed_ms,0,blend_radius_m)
  movel([0.257170, -1.354734, -2.567347, -0.790308, 1.570796, 1.827967],accel_mss,speed_ms,0,blend_radius_m)
  movel([0.257354, -1.354683, -2.567382, -0.790324, 1.570796, 1.828150],accel_mss,speed_ms,0,blend_radius_m)
  movel([0.257671, -1.354609, -2.567432, -0.790348, 1.570796, 1.828467],accel_mss,speed_ms,0,blend_radius_m)
  movel([0.257983, -1.354548, -2.567473, -0.790368, 1.570796, 1.828780],accel_mss,speed_ms,0,blend_radius_m)
  movel([0.258603, -1.354449, -2.567540, -0.790400, 1.570796, 1.829399],accel_mss,speed_ms,0,blend_radius_m)
  movel([0.259219, -1.354355, -2.567603, -0.790430, 1.570796, 1.830015],accel_mss,speed_ms,0,blend_radius_m)
  movel([0.259838, -1.354266, -2.567664, -0.790459, 1.570796, 1.830635],accel_mss,speed_ms,0,blend_radius_m)
  movel([0.260456, -1.354183, -2.567720, -0.790486, 1.570796, 1.831252],accel_mss,speed_ms,0,blend_radius_m)
  movel([0.260762, -1.354149, -2.567743, -0.790497, 1.570796, 1.831558],accel_mss,speed_ms,0,blend_radius_m)
  movel([0.261062, -1.354134, -2.567753, -0.790502, 1.570796, 1.831858],accel_mss,speed_ms,0,blend_radius_m)
  movel([0.261231, -1.354133, -2.567754, -0.790502, 1.570796, 1.832027],accel_mss,speed_ms,0,blend_radius_m)
  movel([0.261397, -1.354144, -2.567746, -0.790499, 1.570796, 1.832193],accel_mss,speed_ms,0,blend_radius_m)
  movel([0.261559, -1.354160, -2.567735, -0.790494, 1.570796, 1.832356],accel_mss,speed_ms,0,blend_radius_m)
  movel([0.261915, -1.354214, -2.567699, -0.790476, 1.570796, 1.832711],accel_mss,speed_ms,0,blend_radius_m)
  movel([0.262265, -1.354278, -2.567656, -0.790455, 1.570796, 1.833062],accel_mss,speed_ms,0,blend_radius_m)
  movel([0.262645, -1.354362, -2.567599, -0.790428, 1.570796, 1.833441],accel_mss,speed_ms,0,blend_radius_m)
  movel([0.263015, -1.354463, -2.567531, -0.790395, 1.570796, 1.833812],accel_mss,speed_ms,0,blend_radius_m)
  movel([0.263373, -1.354584, -2.567449, -0.790356, 1.570796, 1.834169],accel_mss,speed_ms,0,blend_radius_m)
  movel([0.263719, -1.354717, -2.567359, -0.790313, 1.570796, 1.834516],accel_mss,speed_ms,0,blend_radius_m)
  movel([0.264051, -1.354871, -2.567255, -0.790264, 1.570796, 1.834847],accel_mss,speed_ms,0,blend_radius_m)
  movel([0.264368, -1.355040, -2.567140, -0.790209, 1.570796, 1.835164],accel_mss,speed_ms,0,blend_radius_m)
  movel([0.264672, -1.355224, -2.567016, -0.790149, 1.570796, 1.835468],accel_mss,speed_ms,0,blend_radius_m)
  movel([0.264961, -1.355423, -2.566881, -0.790085, 1.570796, 1.835757],accel_mss,speed_ms,0,blend_radius_m)
  movel([0.265237, -1.355638, -2.566735, -0.790016, 1.570796, 1.836033],accel_mss,speed_ms,0,blend_radius_m)
  movel([0.265497, -1.355873, -2.566576, -0.789940, 1.570796, 1.836293],accel_mss,speed_ms,0,blend_radius_m)
  movel([0.265745, -1.356118, -2.566410, -0.789861, 1.570796, 1.836541],accel_mss,speed_ms,0,blend_radius_m)
  movel([0.265974, -1.356379, -2.566232, -0.789777, 1.570796, 1.836770],accel_mss,speed_ms,0,blend_radius_m)
  movel([0.266190, -1.356654, -2.566046, -0.789689, 1.570796, 1.836986],accel_mss,speed_ms,0,blend_radius_m)
  movel([0.266387, -1.356941, -2.565851, -0.789597, 1.570796, 1.837184],accel_mss,speed_ms,0,blend_radius_m)
  movel([0.266567, -1.357243, -2.565646, -0.789501, 1.570796, 1.837363],accel_mss,speed_ms,0,blend_radius_m)
  movel([0.266729, -1.357553, -2.565435, -0.789401, 1.570796, 1.837526],accel_mss,speed_ms,0,blend_radius_m)
  movel([0.266876, -1.357876, -2.565215, -0.789298, 1.570796, 1.837673],accel_mss,speed_ms,0,blend_radius_m)
  movel([0.267004, -1.358211, -2.564987, -0.789191, 1.570796, 1.837800],accel_mss,speed_ms,0,blend_radius_m)
  movel([0.267115, -1.358561, -2.564748, -0.789080, 1.570796, 1.837911],accel_mss,speed_ms,0,blend_radius_m)
  movel([0.267211, -1.358922, -2.564502, -0.788965, 1.570796, 1.838007],accel_mss,speed_ms,0,blend_radius_m)
  movel([0.267286, -1.359290, -2.564251, -0.788848, 1.570796, 1.838082],accel_mss,speed_ms,0,blend_radius_m)
  movel([0.267344, -1.359669, -2.563992, -0.788728, 1.570796, 1.838140],accel_mss,speed_ms,0,blend_radius_m)
  movel([0.267383, -1.360055, -2.563728, -0.788606, 1.570796, 1.838180],accel_mss,speed_ms,0,blend_radius_m)
  movel([0.267406, -1.360450, -2.563458, -0.788481, 1.570796, 1.838202],accel_mss,speed_ms,0,blend_radius_m)
  movel([0.267409, -1.360849, -2.563185, -0.788355, 1.570796, 1.838205],accel_mss,speed_ms,0,blend_radius_m)
  movel([0.267395, -1.361257, -2.562905, -0.788227, 1.570796, 1.838191],accel_mss,speed_ms,0,blend_radius_m)
  movel([0.267361, -1.361670, -2.562622, -0.788097, 1.570796, 1.838158],accel_mss,speed_ms,0,blend_radius_m)
  movel([0.267311, -1.362091, -2.562333, -0.787965, 1.570796, 1.838107],accel_mss,speed_ms,0,blend_radius_m)
  movel([0.267242, -1.362519, -2.562039, -0.787831, 1.570796, 1.838039],accel_mss,speed_ms,0,blend_radius_m)
  movel([0.267157, -1.362949, -2.561744, -0.787697, 1.570796, 1.837953],accel_mss,speed_ms,0,blend_radius_m)
  movel([0.267051, -1.363384, -2.561444, -0.787561, 1.570796, 1.837848],accel_mss,speed_ms,0,blend_radius_m)
  movel([0.266932, -1.363820, -2.561144, -0.787425, 1.570796, 1.837728],accel_mss,speed_ms,0,blend_radius_m)
  movel([0.266795, -1.364258, -2.560842, -0.787289, 1.570796, 1.837591],accel_mss,speed_ms,0,blend_radius_m)
  movel([0.266639, -1.364699, -2.560538, -0.787152, 1.570796, 1.837436],accel_mss,speed_ms,0,blend_radius_m)
  movel([0.266469, -1.365142, -2.560232, -0.787015, 1.570796, 1.837265],accel_mss,speed_ms,0,blend_radius_m)
  movel([0.266281, -1.365582, -2.559928, -0.786879, 1.570796, 1.837077],accel_mss,speed_ms,0,blend_radius_m)
  movel([0.266066, -1.366052, -2.559603, -0.786735, 1.570796, 1.836862],accel_mss,speed_ms,0,blend_radius_m)
  movel([0.265831, -1.366520, -2.559279, -0.786591, 1.570796, 1.836627],accel_mss,speed_ms,0,blend_radius_m)
  movel([0.265580, -1.366985, -2.558956, -0.786448, 1.570796, 1.836377],accel_mss,speed_ms,0,blend_radius_m)
  movel([0.265312, -1.367448, -2.558635, -0.786306, 1.570796, 1.836109],accel_mss,speed_ms,0,blend_radius_m)
  movel([0.265026, -1.367909, -2.558315, -0.786165, 1.570796, 1.835823],accel_mss,speed_ms,0,blend_radius_m)
  movel([0.264726, -1.368365, -2.557998, -0.786026, 1.570796, 1.835522],accel_mss,speed_ms,0,blend_radius_m)
  speed_ms = 0.003
  movel([0.264726, -1.371517, -2.559521, -0.781352, 1.570796, 1.835522],accel_mss,speed_ms,0,blend_radius_m)
  speed_ms = 0.007
  movel([0.264459, -1.371895, -2.559256, -0.781238, 1.570796, 1.835255],accel_mss,speed_ms,0,blend_radius_m)
  movel([0.264181, -1.372273, -2.558992, -0.781124, 1.570796, 1.834978],accel_mss,speed_ms,0,blend_radius_m)
  movel([0.263892, -1.372644, -2.558732, -0.781013, 1.570796, 1.834688],accel_mss,speed_ms,0,blend_radius_m)
  movel([0.263592, -1.373012, -2.558475, -0.780903, 1.570796, 1.834388],accel_mss,speed_ms,0,blend_radius_m)
  movel([0.263283, -1.373372, -2.558222, -0.780795, 1.570796, 1.834079],accel_mss,speed_ms,0,blend_radius_m)
  movel([0.262963, -1.373729, -2.557972, -0.780688, 1.570796, 1.833759],accel_mss,speed_ms,0,blend_radius_m)
  movel([0.262632, -1.374079, -2.557726, -0.780584, 1.570796, 1.833428],accel_mss,speed_ms,0,blend_radius_m)
  movel([0.262300, -1.374415, -2.557490, -0.780484, 1.570796, 1.833096],accel_mss,speed_ms,0,blend_radius_m)
  movel([0.261959, -1.374745, -2.557258, -0.780386, 1.570796, 1.832755],accel_mss,speed_ms,0,blend_radius_m)
  movel([0.261608, -1.375067, -2.557032, -0.780290, 1.570796, 1.832404],accel_mss,speed_ms,0,blend_radius_m)
  movel([0.261251, -1.375381, -2.556810, -0.780197, 1.570796, 1.832047],accel_mss,speed_ms,0,blend_radius_m)
  movel([0.260885, -1.375688, -2.556594, -0.780107, 1.570796, 1.831681],accel_mss,speed_ms,0,blend_radius_m)
  movel([0.260512, -1.375985, -2.556385, -0.780019, 1.570796, 1.831308],accel_mss,speed_ms,0,blend_radius_m)
  movel([0.260133, -1.376274, -2.556181, -0.779934, 1.570796, 1.830929],accel_mss,speed_ms,0,blend_radius_m)
  movel([0.259752, -1.376551, -2.555986, -0.779852, 1.570796, 1.830549],accel_mss,speed_ms,0,blend_radius_m)
  movel([0.259369, -1.376814, -2.555800, -0.779775, 1.570796, 1.830165],accel_mss,speed_ms,0,blend_radius_m)
  movel([0.258979, -1.377071, -2.555619, -0.779699, 1.570796, 1.829775],accel_mss,speed_ms,0,blend_radius_m)
  movel([0.258583, -1.377315, -2.555446, -0.779628, 1.570796, 1.829379],accel_mss,speed_ms,0,blend_radius_m)
  movel([0.258183, -1.377549, -2.555281, -0.779559, 1.570796, 1.828979],accel_mss,speed_ms,0,blend_radius_m)
  movel([0.257780, -1.377770, -2.555124, -0.779494, 1.570796, 1.828576],accel_mss,speed_ms,0,blend_radius_m)
  movel([0.257376, -1.377982, -2.554975, -0.779432, 1.570796, 1.828172],accel_mss,speed_ms,0,blend_radius_m)
  movel([0.256961, -1.378181, -2.554834, -0.779374, 1.570796, 1.827757],accel_mss,speed_ms,0,blend_radius_m)
  movel([0.256546, -1.378366, -2.554703, -0.779320, 1.570796, 1.827342],accel_mss,speed_ms,0,blend_radius_m)
  movel([0.256128, -1.378537, -2.554582, -0.779270, 1.570796, 1.826924],accel_mss,speed_ms,0,blend_radius_m)
  movel([0.255708, -1.378690, -2.554473, -0.779226, 1.570796, 1.826504],accel_mss,speed_ms,0,blend_radius_m)
  movel([0.255290, -1.378829, -2.554375, -0.779185, 1.570796, 1.826086],accel_mss,speed_ms,0,blend_radius_m)
  movel([0.254850, -1.378958, -2.554283, -0.779148, 1.570796, 1.825646],accel_mss,speed_ms,0,blend_radius_m)
  movel([0.254411, -1.379071, -2.554203, -0.779115, 1.570796, 1.825208],accel_mss,speed_ms,0,blend_radius_m)
  movel([0.253975, -1.379170, -2.554133, -0.779086, 1.570796, 1.824771],accel_mss,speed_ms,0,blend_radius_m)
  movel([0.253540, -1.379256, -2.554072, -0.779061, 1.570796, 1.824336],accel_mss,speed_ms,0,blend_radius_m)
  movel([0.253112, -1.379324, -2.554024, -0.779041, 1.570796, 1.823908],accel_mss,speed_ms,0,blend_radius_m)
  movel([0.252686, -1.379377, -2.553986, -0.779026, 1.570796, 1.823483],accel_mss,speed_ms,0,blend_radius_m)
  movel([0.252264, -1.379416, -2.553958, -0.779015, 1.570796, 1.823061],accel_mss,speed_ms,0,blend_radius_m)
  movel([0.251849, -1.379438, -2.553943, -0.779008, 1.570796, 1.822646],accel_mss,speed_ms,0,blend_radius_m)
  movel([0.251441, -1.379446, -2.553937, -0.779006, 1.570796, 1.822237],accel_mss,speed_ms,0,blend_radius_m)
  movel([0.251039, -1.379436, -2.553944, -0.779009, 1.570796, 1.821835],accel_mss,speed_ms,0,blend_radius_m)
  movel([0.250665, -1.379411, -2.553962, -0.779016, 1.570796, 1.821461],accel_mss,speed_ms,0,blend_radius_m)
  movel([0.250299, -1.379371, -2.553991, -0.779028, 1.570796, 1.821095],accel_mss,speed_ms,0,blend_radius_m)
  movel([0.249945, -1.379311, -2.554033, -0.779045, 1.570796, 1.820742],accel_mss,speed_ms,0,blend_radius_m)
  movel([0.249601, -1.379236, -2.554086, -0.779067, 1.570796, 1.820397],accel_mss,speed_ms,0,blend_radius_m)
  movel([0.249268, -1.379142, -2.554153, -0.779094, 1.570796, 1.820064],accel_mss,speed_ms,0,blend_radius_m)
  movel([0.248923, -1.379026, -2.554235, -0.779128, 1.570796, 1.819719],accel_mss,speed_ms,0,blend_radius_m)
  movel([0.248591, -1.378894, -2.554329, -0.779166, 1.570796, 1.819387],accel_mss,speed_ms,0,blend_radius_m)
  movel([0.248271, -1.378745, -2.554435, -0.779210, 1.570796, 1.819067],accel_mss,speed_ms,0,blend_radius_m)
  movel([0.247963, -1.378581, -2.554551, -0.779258, 1.570796, 1.818760],accel_mss,speed_ms,0,blend_radius_m)
  movel([0.247671, -1.378402, -2.554677, -0.779310, 1.570796, 1.818468],accel_mss,speed_ms,0,blend_radius_m)
  movel([0.247393, -1.378209, -2.554814, -0.779366, 1.570796, 1.818189],accel_mss,speed_ms,0,blend_radius_m)
  movel([0.247127, -1.378000, -2.554962, -0.779427, 1.570796, 1.817923],accel_mss,speed_ms,0,blend_radius_m)
  movel([0.246876, -1.377779, -2.555118, -0.779492, 1.570796, 1.817673],accel_mss,speed_ms,0,blend_radius_m)
  movel([0.246644, -1.377540, -2.555287, -0.779562, 1.570796, 1.817440],accel_mss,speed_ms,0,blend_radius_m)
  movel([0.246416, -1.377284, -2.555468, -0.779637, 1.570796, 1.817213],accel_mss,speed_ms,0,blend_radius_m)
  movel([0.246206, -1.377014, -2.555659, -0.779716, 1.570796, 1.817002],accel_mss,speed_ms,0,blend_radius_m)
  movel([0.246010, -1.376733, -2.555857, -0.779799, 1.570796, 1.816806],accel_mss,speed_ms,0,blend_radius_m)
  movel([0.245831, -1.376439, -2.556065, -0.779885, 1.570796, 1.816628],accel_mss,speed_ms,0,blend_radius_m)
  movel([0.245667, -1.376134, -2.556280, -0.779975, 1.570796, 1.816463],accel_mss,speed_ms,0,blend_radius_m)
  movel([0.245521, -1.375818, -2.556503, -0.780068, 1.570796, 1.816318],accel_mss,speed_ms,0,blend_radius_m)
  movel([0.245390, -1.375493, -2.556732, -0.780164, 1.570796, 1.816186],accel_mss,speed_ms,0,blend_radius_m)
  movel([0.245275, -1.375156, -2.556969, -0.780264, 1.570796, 1.816071],accel_mss,speed_ms,0,blend_radius_m)
  movel([0.245179, -1.374811, -2.557212, -0.780367, 1.570796, 1.815975],accel_mss,speed_ms,0,blend_radius_m)
  movel([0.245098, -1.374449, -2.557466, -0.780474, 1.570796, 1.815894],accel_mss,speed_ms,0,blend_radius_m)
  movel([0.245033, -1.374081, -2.557724, -0.780583, 1.570796, 1.815829],accel_mss,speed_ms,0,blend_radius_m)
  movel([0.244986, -1.373704, -2.557989, -0.780696, 1.570796, 1.815783],accel_mss,speed_ms,0,blend_radius_m)
  movel([0.244956, -1.373320, -2.558259, -0.780811, 1.570796, 1.815752],accel_mss,speed_ms,0,blend_radius_m)
  movel([0.244943, -1.372928, -2.558533, -0.780928, 1.570796, 1.815739],accel_mss,speed_ms,0,blend_radius_m)
  movel([0.244948, -1.372529, -2.558813, -0.781047, 1.570796, 1.815745],accel_mss,speed_ms,0,blend_radius_m)
  movel([0.244971, -1.372125, -2.559095, -0.781169, 1.570796, 1.815768],accel_mss,speed_ms,0,blend_radius_m)
  movel([0.245012, -1.371714, -2.559383, -0.781292, 1.570796, 1.815809],accel_mss,speed_ms,0,blend_radius_m)
  movel([0.245068, -1.371300, -2.559672, -0.781417, 1.570796, 1.815864],accel_mss,speed_ms,0,blend_radius_m)
  movel([0.245143, -1.370883, -2.559963, -0.781543, 1.570796, 1.815940],accel_mss,speed_ms,0,blend_radius_m)
  movel([0.245235, -1.370463, -2.560256, -0.781670, 1.570796, 1.816032],accel_mss,speed_ms,0,blend_radius_m)
  movel([0.245345, -1.370040, -2.560551, -0.781798, 1.570796, 1.816141],accel_mss,speed_ms,0,blend_radius_m)
  movel([0.245471, -1.369612, -2.560849, -0.781928, 1.570796, 1.816268],accel_mss,speed_ms,0,blend_radius_m)
  movel([0.245615, -1.369183, -2.561147, -0.782059, 1.570796, 1.816411],accel_mss,speed_ms,0,blend_radius_m)
  movel([0.245777, -1.368753, -2.561446, -0.782190, 1.570796, 1.816573],accel_mss,speed_ms,0,blend_radius_m)
  movel([0.245954, -1.368323, -2.561744, -0.782321, 1.570796, 1.816750],accel_mss,speed_ms,0,blend_radius_m)
  movel([0.246150, -1.367890, -2.562045, -0.782454, 1.570796, 1.816946],accel_mss,speed_ms,0,blend_radius_m)
  movel([0.246359, -1.367459, -2.562344, -0.782586, 1.570796, 1.817156],accel_mss,speed_ms,0,blend_radius_m)
  movel([0.246577, -1.367041, -2.562633, -0.782715, 1.570796, 1.817373],accel_mss,speed_ms,0,blend_radius_m)
  movel([0.246806, -1.366624, -2.562922, -0.782843, 1.570796, 1.817603],accel_mss,speed_ms,0,blend_radius_m)
  movel([0.247047, -1.366208, -2.563209, -0.782971, 1.570796, 1.817843],accel_mss,speed_ms,0,blend_radius_m)
  movel([0.247299, -1.365793, -2.563496, -0.783100, 1.570796, 1.818095],accel_mss,speed_ms,0,blend_radius_m)
  movel([0.247538, -1.365421, -2.563753, -0.783215, 1.570796, 1.818334],accel_mss,speed_ms,0,blend_radius_m)
  movel([0.247791, -1.365054, -2.564006, -0.783329, 1.570796, 1.818588],accel_mss,speed_ms,0,blend_radius_m)
  movel([0.248054, -1.364689, -2.564258, -0.783442, 1.570796, 1.818850],accel_mss,speed_ms,0,blend_radius_m)
  movel([0.248331, -1.364330, -2.564505, -0.783554, 1.570796, 1.819128],accel_mss,speed_ms,0,blend_radius_m)
  movel([0.248616, -1.363978, -2.564747, -0.783663, 1.570796, 1.819412],accel_mss,speed_ms,0,blend_radius_m)
  movel([0.248911, -1.363632, -2.564986, -0.783772, 1.570796, 1.819708],accel_mss,speed_ms,0,blend_radius_m)
  movel([0.249219, -1.363292, -2.565219, -0.783878, 1.570796, 1.820015],accel_mss,speed_ms,0,blend_radius_m)
  movel([0.249537, -1.362959, -2.565448, -0.783982, 1.570796, 1.820333],accel_mss,speed_ms,0,blend_radius_m)
  movel([0.249891, -1.362605, -2.565691, -0.784093, 1.570796, 1.820687],accel_mss,speed_ms,0,blend_radius_m)
  movel([0.250253, -1.362257, -2.565930, -0.784203, 1.570796, 1.821049],accel_mss,speed_ms,0,blend_radius_m)
  movel([0.250622, -1.361915, -2.566164, -0.784310, 1.570796, 1.821419],accel_mss,speed_ms,0,blend_radius_m)
  movel([0.251000, -1.361582, -2.566392, -0.784415, 1.570796, 1.821796],accel_mss,speed_ms,0,blend_radius_m)
  movel([0.251409, -1.361232, -2.566632, -0.784525, 1.570796, 1.822206],accel_mss,speed_ms,0,blend_radius_m)
  movel([0.251825, -1.360894, -2.566863, -0.784632, 1.570796, 1.822622],accel_mss,speed_ms,0,blend_radius_m)
  movel([0.252250, -1.360562, -2.567090, -0.784737, 1.570796, 1.823046],accel_mss,speed_ms,0,blend_radius_m)
  movel([0.252636, -1.360275, -2.567286, -0.784828, 1.570796, 1.823432],accel_mss,speed_ms,0,blend_radius_m)
  movel([0.253029, -1.359998, -2.567475, -0.784916, 1.570796, 1.823825],accel_mss,speed_ms,0,blend_radius_m)
  movel([0.253428, -1.359732, -2.567656, -0.785000, 1.570796, 1.824225],accel_mss,speed_ms,0,blend_radius_m)
  movel([0.253830, -1.359485, -2.567825, -0.785079, 1.570796, 1.824626],accel_mss,speed_ms,0,blend_radius_m)
  movel([0.254233, -1.359250, -2.567985, -0.785154, 1.570796, 1.825029],accel_mss,speed_ms,0,blend_radius_m)
  movel([0.254642, -1.359027, -2.568137, -0.785225, 1.570796, 1.825438],accel_mss,speed_ms,0,blend_radius_m)
  movel([0.255090, -1.358801, -2.568291, -0.785297, 1.570796, 1.825886],accel_mss,speed_ms,0,blend_radius_m)
  movel([0.255537, -1.358586, -2.568437, -0.785366, 1.570796, 1.826333],accel_mss,speed_ms,0,blend_radius_m)
  movel([0.255988, -1.358384, -2.568575, -0.785430, 1.570796, 1.826784],accel_mss,speed_ms,0,blend_radius_m)
  movel([0.256396, -1.358210, -2.568693, -0.785486, 1.570796, 1.827192],accel_mss,speed_ms,0,blend_radius_m)
  movel([0.256803, -1.358048, -2.568804, -0.785538, 1.570796, 1.827599],accel_mss,speed_ms,0,blend_radius_m)
  movel([0.256987, -1.357978, -2.568851, -0.785560, 1.570796, 1.827783],accel_mss,speed_ms,0,blend_radius_m)
  movel([0.257170, -1.357918, -2.568892, -0.785579, 1.570796, 1.827967],accel_mss,speed_ms,0,blend_radius_m)
  movel([0.257354, -1.357866, -2.568927, -0.785596, 1.570796, 1.828150],accel_mss,speed_ms,0,blend_radius_m)
  movel([0.257671, -1.357792, -2.568977, -0.785620, 1.570796, 1.828467],accel_mss,speed_ms,0,blend_radius_m)
  movel([0.257983, -1.357732, -2.569018, -0.785639, 1.570796, 1.828780],accel_mss,speed_ms,0,blend_radius_m)
  movel([0.258603, -1.357633, -2.569085, -0.785671, 1.570796, 1.829399],accel_mss,speed_ms,0,blend_radius_m)
  movel([0.259219, -1.357539, -2.569149, -0.785701, 1.570796, 1.830015],accel_mss,speed_ms,0,blend_radius_m)
  movel([0.259838, -1.357450, -2.569210, -0.785729, 1.570796, 1.830635],accel_mss,speed_ms,0,blend_radius_m)
  movel([0.260456, -1.357367, -2.569266, -0.785756, 1.570796, 1.831252],accel_mss,speed_ms,0,blend_radius_m)
  movel([0.260762, -1.357333, -2.569289, -0.785767, 1.570796, 1.831558],accel_mss,speed_ms,0,blend_radius_m)
  movel([0.261062, -1.357318, -2.569299, -0.785772, 1.570796, 1.831858],accel_mss,speed_ms,0,blend_radius_m)
  movel([0.261231, -1.357317, -2.569300, -0.785772, 1.570796, 1.832027],accel_mss,speed_ms,0,blend_radius_m)
  movel([0.261397, -1.357328, -2.569292, -0.785768, 1.570796, 1.832193],accel_mss,speed_ms,0,blend_radius_m)
  movel([0.261559, -1.357344, -2.569281, -0.785763, 1.570796, 1.832356],accel_mss,speed_ms,0,blend_radius_m)
  movel([0.261915, -1.357398, -2.569245, -0.785746, 1.570796, 1.832711],accel_mss,speed_ms,0,blend_radius_m)
  movel([0.262265, -1.357462, -2.569201, -0.785725, 1.570796, 1.833062],accel_mss,speed_ms,0,blend_radius_m)
  movel([0.262645, -1.357546, -2.569145, -0.785699, 1.570796, 1.833441],accel_mss,speed_ms,0,blend_radius_m)
  movel([0.263015, -1.357647, -2.569076, -0.785666, 1.570796, 1.833812],accel_mss,speed_ms,0,blend_radius_m)
  movel([0.263373, -1.357767, -2.568994, -0.785628, 1.570796, 1.834169],accel_mss,speed_ms,0,blend_radius_m)
  movel([0.263719, -1.357900, -2.568904, -0.785585, 1.570796, 1.834516],accel_mss,speed_ms,0,blend_radius_m)
  movel([0.264051, -1.358053, -2.568800, -0.785536, 1.570796, 1.834847],accel_mss,speed_ms,0,blend_radius_m)
  movel([0.264368, -1.358222, -2.568685, -0.785482, 1.570796, 1.835164],accel_mss,speed_ms,0,blend_radius_m)
  movel([0.264672, -1.358406, -2.568560, -0.785423, 1.570796, 1.835468],accel_mss,speed_ms,0,blend_radius_m)
  movel([0.264961, -1.358605, -2.568425, -0.785360, 1.570796, 1.835757],accel_mss,speed_ms,0,blend_radius_m)
  movel([0.265237, -1.358819, -2.568279, -0.785291, 1.570796, 1.836033],accel_mss,speed_ms,0,blend_radius_m)
  movel([0.265497, -1.359053, -2.568119, -0.785217, 1.570796, 1.836293],accel_mss,speed_ms,0,blend_radius_m)
  movel([0.265745, -1.359298, -2.567952, -0.785139, 1.570796, 1.836541],accel_mss,speed_ms,0,blend_radius_m)
  movel([0.265974, -1.359559, -2.567775, -0.785056, 1.570796, 1.836770],accel_mss,speed_ms,0,blend_radius_m)
  movel([0.266190, -1.359832, -2.567588, -0.784969, 1.570796, 1.836986],accel_mss,speed_ms,0,blend_radius_m)
  movel([0.266387, -1.360119, -2.567392, -0.784878, 1.570796, 1.837184],accel_mss,speed_ms,0,blend_radius_m)
  movel([0.266567, -1.360420, -2.567187, -0.784782, 1.570796, 1.837363],accel_mss,speed_ms,0,blend_radius_m)
  movel([0.266729, -1.360729, -2.566975, -0.784684, 1.570796, 1.837526],accel_mss,speed_ms,0,blend_radius_m)
  movel([0.266876, -1.361052, -2.566755, -0.784582, 1.570796, 1.837673],accel_mss,speed_ms,0,blend_radius_m)
  movel([0.267004, -1.361386, -2.566526, -0.784477, 1.570796, 1.837800],accel_mss,speed_ms,0,blend_radius_m)
  movel([0.267115, -1.361735, -2.566287, -0.784367, 1.570796, 1.837911],accel_mss,speed_ms,0,blend_radius_m)
  movel([0.267211, -1.362095, -2.566040, -0.784253, 1.570796, 1.838007],accel_mss,speed_ms,0,blend_radius_m)
  movel([0.267286, -1.362462, -2.565789, -0.784138, 1.570796, 1.838082],accel_mss,speed_ms,0,blend_radius_m)
  movel([0.267344, -1.362841, -2.565529, -0.784019, 1.570796, 1.838140],accel_mss,speed_ms,0,blend_radius_m)
  movel([0.267383, -1.363226, -2.565265, -0.783899, 1.570796, 1.838180],accel_mss,speed_ms,0,blend_radius_m)
  movel([0.267406, -1.363619, -2.564994, -0.783776, 1.570796, 1.838202],accel_mss,speed_ms,0,blend_radius_m)
  movel([0.267409, -1.364018, -2.564720, -0.783651, 1.570796, 1.838205],accel_mss,speed_ms,0,blend_radius_m)
  movel([0.267395, -1.364425, -2.564440, -0.783524, 1.570796, 1.838191],accel_mss,speed_ms,0,blend_radius_m)
  movel([0.267361, -1.364837, -2.564156, -0.783396, 1.570796, 1.838158],accel_mss,speed_ms,0,blend_radius_m)
  movel([0.267311, -1.365257, -2.563866, -0.783266, 1.570796, 1.838107],accel_mss,speed_ms,0,blend_radius_m)
  movel([0.267242, -1.365684, -2.563572, -0.783134, 1.570796, 1.838039],accel_mss,speed_ms,0,blend_radius_m)
  movel([0.267157, -1.366113, -2.563275, -0.783001, 1.570796, 1.837953],accel_mss,speed_ms,0,blend_radius_m)
  movel([0.267051, -1.366546, -2.562976, -0.782867, 1.570796, 1.837848],accel_mss,speed_ms,0,blend_radius_m)
  movel([0.266932, -1.366982, -2.562674, -0.782733, 1.570796, 1.837728],accel_mss,speed_ms,0,blend_radius_m)
  movel([0.266795, -1.367419, -2.562371, -0.782598, 1.570796, 1.837591],accel_mss,speed_ms,0,blend_radius_m)
  movel([0.266639, -1.367859, -2.562067, -0.782463, 1.570796, 1.837436],accel_mss,speed_ms,0,blend_radius_m)
  movel([0.266469, -1.368300, -2.561760, -0.782328, 1.570796, 1.837265],accel_mss,speed_ms,0,blend_radius_m)
  movel([0.266281, -1.368740, -2.561455, -0.782194, 1.570796, 1.837077],accel_mss,speed_ms,0,blend_radius_m)
  movel([0.266066, -1.369208, -2.561129, -0.782051, 1.570796, 1.836862],accel_mss,speed_ms,0,blend_radius_m)
  movel([0.265831, -1.369675, -2.560805, -0.781909, 1.570796, 1.836627],accel_mss,speed_ms,0,blend_radius_m)
  movel([0.265580, -1.370140, -2.560481, -0.781768, 1.570796, 1.836377],accel_mss,speed_ms,0,blend_radius_m)
  movel([0.265312, -1.370602, -2.560159, -0.781628, 1.570796, 1.836109],accel_mss,speed_ms,0,blend_radius_m)
  movel([0.265026, -1.371061, -2.559838, -0.781489, 1.570796, 1.835823],accel_mss,speed_ms,0,blend_radius_m)
  movel([0.264726, -1.371517, -2.559521, -0.781352, 1.570796, 1.835522],accel_mss,speed_ms,0,blend_radius_m)
  speed_ms = 0.003
  movel([0.264726, -1.359043, -2.553380, -0.799966, 1.570796, 1.835522],accel_mss,speed_ms,0,blend_radius_m)
  speed_ms = 0.01
  movel([0.264726, -1.335140, -2.540718, -0.836531, 1.570796, 1.835522],accel_mss,speed_ms,0,blend_radius_m)
  movel([0.175631, -1.289895, -2.569395, -0.853098, 1.570796, 1.746427],accel_mss,speed_ms,0,blend_radius_m)
  movel([0.175631, -1.235022, -2.534278, -0.943089, 1.570796, 1.746427],accel_mss,speed_ms,0,blend_radius_m)
  # End of main program
end

Machining2()=
